(* IEC 61131-3 sources: Antarbhukti-LLM/DatasetCreation/SeedSTs/batch2_filtered_NETWORK (part 2) *)

(* ---- HTTP_GET.ST ---- *)
(*@PROPERTIES_EX@
TYPE: POU
LOCALE: 0
IEC_LANGUAGE: ST
PLC_TYPE: independent
PROC_TYPE: independent
GROUP: NETWORK
*)
(*@KEY@:DESCRIPTION*)

version 1.3	12. apr. 2011
programmer 	ks
tested by	ks

HTTP_GET führt eine HTTP Abfrage einer Web-Seite bei einem WEB_Server durch, und stellt die Daten ausbereitet zu verfügung
(*@KEY@:END_DESCRIPTION*)
FUNCTION_BLOCK HTTP_GET

(*Group:Default*)

VAR_IN_OUT
	URL_DATA :	oscat_url;
	IP_C :	oscat_IP_C;(*IP_Control Verwaltungsstruktur*)
	S_BUF :	oscat_NETWORK_BUFFER;
	R_BUF :	oscat_NETWORK_BUFFER;
END_VAR

VAR_INPUT
	IP4 :	DWORD;
	GET :	BOOL;
	MODE :	BYTE := BYTE#2;
	UNLOCK_BUF :	BOOL;
END_VAR

VAR_OUTPUT
	HTTP_STATUS :	STRING;
	HEADER_START :	UINT;(*HTTP Header (Message Header)*)
	HEADER_STOP :	UINT;(*HTTP Header (Message Header)*)
	BODY_START :	UINT;(*Message Body*)
	BODY_STOP :	UINT;(*Message Body*)
	DONE :	BOOL;
	ERROR :	DWORD;
END_VAR

VAR
	READ_HTTP :	READ_HTTP;
	BUFFER_SEARCH :	BUFFER_SEARCH_NW;
	_STRING_TO_BUFFER :	_STRING_TO_BUFFER_NW;
	IP_FIFO :	IP_FIFO;
	IS_NUM :	IS_NUM;
	ip_state :	BYTE;
	ip_id :	BYTE;
	get_last :	BOOL;
	ip4_stored :	DWORD;
	state :	INT;
	i :	INT;
	http_1_1_host :	BOOL;
	total_size :	INT;
	text :	oscat_STRING250;
	delimiter2b :	oscat_STRING2;
	delimiter4b :	oscat_STRING4;
	del_end :	oscat_STRING4;
	del_pos :	INT;
	idx :	INT;
	rcv_timeout :	BOOL;
	con_rdce :	BOOL;
END_VAR

(*Group:debug*)

VAR
	(*<LOG_MSG :	LOG_MSG;>*)
END_VAR

VAR_EXTERNAL
	(*<LOG_CL :	us_LOG_CONTROL;>*)(*Debug-Datenstruktur*)
END_VAR

VAR
	(*<_debug_enable :	BOOL := TRUE;>*)
END_VAR

(*@KEY@: WORKSHEET
NAME: HTTP_GET
IEC_LANGUAGE: ST
*)

CASE state OF
00:	IF GET AND NOT get_last THEN (* auf positive Flanke SET warten *)
		state        := 10;
		ip4_stored   := IP4; (* aktuelle IP4 speichern *)
		DONE         := FALSE;
		total_size   := 0;
		HEADER_START := UINT#0;
		HEADER_STOP  := UINT#0;
		BODY_START   := UINT#0;
		BODY_STOP    := UINT#0;
		HTTP_STATUS  := '';
    	ERROR        := DWORD#0;
    	ip_state     := BYTE#1; (* Anmelden *)

    	(* workaround für pcworx -> kein $0D$0A als Stringkonstante möglich *)
    	delimiter2b := CONCAT(BYTE_TO_STRING(BYTE#16#0D,'%c'),BYTE_TO_STRING(BYTE#16#0A,'%c'));
    	delimiter4b := CONCAT(delimiter2b,delimiter2b);
        (*####################  DEBUG-MESSAGE  ###################################*)
        (*IF _debug_enable THEN
            LOG_CL.NEW_MSG := 'HTTP: S00 START /IP_ID ~4';
            LOG_CL.PRINTF[4]  := BYTE_TO_STRING(IP_ID,'%u');
            LOG_MSG();
        END_IF;*)
        (*########################################################################*)
  	END_IF;

10:	IF ip_state = BYTE#3 THEN (* Bei IP_Control anmelden und auf freigabe warten *)
		idx := 0;
		text := CONCAT('GET ',URL_DATA.PATH);
		_STRING_TO_BUFFER(STR:=text,POS:=idx,PT:=S_BUF.BUFFER,SIZE:=UINT#4096); (* GET path in buffer kopieren *)
		S_BUF.BUFFER:=_STRING_TO_BUFFER.pt;
		idx := idx + LEN(text);

		IF LEN(URL_DATA.QUERY) > 0 THEN
			S_BUF.BUFFER[idx] := BYTE#63; (* ASCII '?' *)
			idx := idx + 1;
			_STRING_TO_BUFFER(STR:=URL_DATA.QUERY,POS:=idx,PT:=S_BUF.BUFFER,SIZE:=UINT#4096); (* QUERY in buffer kopieren *)
			S_BUF.BUFFER:=_STRING_TO_BUFFER.pt;
			idx := idx + LEN(URL_DATA.QUERY);
		END_IF;

		IF MODE >= BYTE#2 THEN (* gewünschte HTTP Version uebergeben *)
			text := ' HTTP/1.1';
		ELSE
			text := ' HTTP/1.0';
		END_IF;
		text := CONCAT(text,delimiter2b);
		_STRING_TO_BUFFER(STR:=text,POS:=idx,PT:=S_BUF.BUFFER,SIZE:=UINT#4096); (* HTTP Version in buffer kopieren *)
		S_BUF.BUFFER:=_STRING_TO_BUFFER.pt;
		idx := idx + LEN(text);

		IF MODE = BYTE#1 THEN (* HTTP/1.0 mit persistenter Verbindung gewünscht *)
			text := CONCAT('Connection: Keep-Alive',delimiter2b); (* workaround für pcworx -> kein $0D$0A als Stringkonstante möglich *)
		ELSIF MODE = BYTE#3 THEN (* HTTP/1.1 ohne persistenter Verbindung gewünscht *)
			text := CONCAT('Connection: Close',delimiter2b); (* workaround für pcworx -> kein $0D$0A als Stringkonstante möglich *)
		ELSE
			text := '';
		END_IF;
		text := CONCAT(text,URL_DATA.HEADER);
		_STRING_TO_BUFFER(STR:=text,POS:=idx,PT:=S_BUF.BUFFER,SIZE:=UINT#4096); (* HTTP Version in buffer kopieren *)
		S_BUF.BUFFER:=_STRING_TO_BUFFER.pt;
		idx := idx + LEN(text);

		text := CONCAT('Host: ',URL_DATA.DOMAIN);
		text := CONCAT(text,delimiter4b); (* workaround für pcworx -> kein $0D$0A als Stringkonstante möglich *)
		_STRING_TO_BUFFER(STR:=text,POS:=idx,PT:=S_BUF.BUFFER,SIZE:=UINT#4096); (* HTTP Host in buffer kopieren *)
		S_BUF.BUFFER:=_STRING_TO_BUFFER.pt;
		idx := idx + LEN(text);

		(* IP Datenverkehr einrichten *)
		IF URL_DATA.PORT = WORD#0 THEN
			IP_C.C_PORT    := WORD#80;        (* Standard-Portnummer verwenden               *)
		ELSE
			IP_C.C_PORT    := URL_DATA.PORT;  (* Portnummer aus URL verwenden                *)
		END_IF;

		IP_C.C_IP       := ip4_stored;       (* IP eintragen                                  *)
		IP_C.C_MODE     := BYTE#0;           (* Mode: TCP+AKTIV+PORT+IP                       *)
		IP_C.C_ENABLE   := TRUE;             (* Verbindungsaufbau freigeben                   *)
		IP_C.TIME_RESET := TRUE;             (* Zeitueberwachung rücksetzen                   *)
		IP_C.R_OBSERVE  := TRUE;             (* Datenempfang ueberwachen                      *)
		S_BUF.SIZE      := INT_TO_UINT(idx); (* Sendelänge eintragen                          *)
		R_BUF.SIZE      := UINT#0;           (* Empfangslänge rücksetzen                      *)

		state := 30;
        (*####################  DEBUG-MESSAGE  ###################################*)
        (*IF _debug_enable THEN
            LOG_CL.NEW_MSG := 'HTTP: S20 SEND /IP_ID ~4';
            LOG_CL.PRINTF[4]  := BYTE_TO_STRING(IP_ID,'%u');
            LOG_MSG();
        END_IF;*)
        (*########################################################################*)

	END_IF;

30:	rcv_timeout := (IP_C.ERROR AND DWORD#16#0000_FF00) = DWORD#16#0000_FF00;
	con_rdce := (IP_C.ERROR AND DWORD#16#FD00_0000) = DWORD#16#FD00_0000;

	IF S_BUF.SIZE = UINT#0 THEN
		IF total_size = 0 THEN
			IF R_BUF.SIZE > UINT#15 THEN;  (* länge der empfangenen Daten prüfen *)

				(* HTTP HEADER Ende suchen -> durch $0D$A$0D$A erkennbar bei DEC RT-11,CP/M,MS-DOS,Windows *)
				del_end := delimiter4b;

				BUFFER_SEARCH(size:=R_BUF.SIZE,str:=del_end,pos:=0,ign:=FALSE,pt:=R_BUF.BUFFER);
				R_BUF.BUFFER:=BUFFER_SEARCH.pt;
				del_pos := BUFFER_SEARCH.BUFFER_SEARCH;

				(* kein Ende gefunden ? -> andere Ende-Codierung suchen *)
				IF del_pos = 0 THEN
          			(* workaround für pcworx -> kein $0A$0A als Stringkonstante möglich *)
          			del_end := CONCAT(BYTE_TO_STRING(BYTE#16#0A,'%c'),BYTE_TO_STRING(BYTE#16#0A,'%c'));

          			(* HTTP HEADER Ende suchen -> durch $A$A erkennbar bei Multics, Unix-Derivate,Mac OS X *)
          			BUFFER_SEARCH(size:=R_BUF.SIZE,str:=del_end,pos:=0,ign:=FALSE,pt:=R_BUF.BUFFER);
          			R_BUF.BUFFER:=BUFFER_SEARCH.pt;
		  			del_pos := BUFFER_SEARCH.BUFFER_SEARCH;
        		END_IF;

				IF del_pos > 0 THEN
					HEADER_START := UINT#0;
					HEADER_STOP  := INT_TO_UINT(del_pos + LEN(del_end) - 1);
					TOTAL_SIZE   := -1; (* HTTP Header empfangen aber noch keine gesamtlänge bekannt *)
				END_IF;

                (*####################  DEBUG-MESSAGE  ###################################*)
                (*IF _debug_enable THEN
                    LOG_CL.NEW_MSG := 'HTTP: S20 HEADER_START ~1 / HEADER_STOP ~2/IP_ID ~4';
                    LOG_CL.PRINTF[4]  := BYTE_TO_STRING(IP_ID,'%u');
                    LOG_CL.PRINTF[1]  := UINT_TO_STRING(HEADER_START,'%u');
                    LOG_CL.PRINTF[2]  := UINT_TO_STRING(HEADER_STOP,'%u');
                    LOG_MSG();
                END_IF;*)
                (*########################################################################*)

				(* HTTP Statuscode auswerten: (kann 1.0 oder 1.1 sein *)
				READ_HTTP(size:=HEADER_STOP,pos:=0,SRC:='',pt:=R_BUF.BUFFER);
				R_BUF.BUFFER:=READ_HTTP.pt;

				i := LEN(READ_HTTP.READ_HTTP);
				IF i > 7 THEN
					(* HTTP Version von HOST auswerten 1.0 oder 1.1 *)
					text:=MID(READ_HTTP.READ_HTTP,1,3);
					http_1_1_host := EQ_STRING(text,'1');

					(* Code und Meldung isolieren *)
					HTTP_STATUS := RIGHT(READ_HTTP.READ_HTTP,i - 4);
				END_IF;

				(* positive HTTP Anfrage ? *)
				IF FIND(HTTP_STATUS,'200') > 0 THEN

					(* 'Content-Length: Wert einlesen auswerten *)
					READ_HTTP(size:=HEADER_STOP,pos:=0,SRC:='CONTENT-LENGTH',pt:=R_BUF.BUFFER);
					R_BUF.BUFFER:=READ_HTTP.pt;
					text:=READ_HTTP.READ_HTTP;

					IF LEN(text) > 0 AND LEN(text) <= 80 THEN
						IS_NUM(str:=text);
						IF IS_NUM.IS_NUM THEN
							(* erwartete gesamtmenge an Bytes berechnen *)
							total_size := STRING_TO_INT(text)+ UINT_TO_INT(HEADER_STOP) + 1;
                            (*####################  DEBUG-MESSAGE  ###################################*)
                            (*IF _debug_enable THEN
                                LOG_CL.NEW_MSG := 'HTTP: S20 HEADER ~1, BODY ~2 TOTAL ~3 /IP_ID ~4';
                                LOG_CL.PRINTF[4]  := BYTE_TO_STRING(IP_ID,'%u');
                                LOG_CL.PRINTF[1]  := UINT_TO_STRING(HEADER_STOP,'%u');
                                LOG_CL.PRINTF[2]  := INT_TO_STRING(TOTAL_SIZE-UINT_TO_INT(HEADER_STOP),'%d');
                                LOG_CL.PRINTF[3]  := INT_TO_STRING(TOTAL_SIZE,'%d');
                                LOG_MSG();
                            END_IF;*)
                            (*########################################################################*)
						END_IF;
					END_IF;
				ELSE
					ERROR := DWORD#16#000000FC; (* Fehler durch HTTP-Statuscodes *)
				END_IF;
			END_IF;
			(* 1. bei bekannter Content-Length wird nach erhalt der erwartenen Daten die verbindung beendet *)
			(* 2. bei persistenter Verbindung muss bei unbekannter Datenmenge auf Receive-Timeout gewartet werden *)
			(* 3. wenn nach datenempfang die verbindung vom host unterbrochen wird *)
		ELSIF (R_BUF.SIZE >= INT_TO_UINT(total_size)) OR
			(R_BUF.SIZE > UINT#0 AND total_size < 0 AND ((rcv_timeout OR con_rdce) OR (IP_C.C_STATE = BYTE#1))) THEN

			IF R_BUF.SIZE - UINT#1 > HEADER_STOP THEN (* BODY Daten vorhanden *)
				BODY_START := HEADER_STOP + UINT#1;
				BODY_STOP  := R_BUF.SIZE - UINT#1;
                (*####################  DEBUG-MESSAGE  ###################################*)
                (*IF _debug_enable THEN
                    LOG_CL.NEW_MSG := 'HTTP: S20 BODY ~1, START ~2 END ~3 /IP_ID ~4';
                    LOG_CL.PRINTF[4]  := BYTE_TO_STRING(IP_ID,'%u');
                    LOG_CL.PRINTF[1]  := UINT_TO_STRING(HEADER_STOP,'%u');
                    LOG_CL.PRINTF[2]  := UINT_TO_STRING(BODY_START,'%u');
                    LOG_CL.PRINTF[3]  := UINT_TO_STRING(BODY_STOP,'%u');
                    LOG_MSG();
                END_IF;*)
                (*########################################################################*)

			END_IF;

			DONE := TRUE;
			IP_C.C_ENABLE := FALSE; (* Verbindung abbauen  *)
			state := 40;
            (*####################  DEBUG-MESSAGE  ###################################*)
            (*IF _debug_enable THEN
                LOG_CL.NEW_MSG := 'HTTP: S30 OK /IP_ID ~4';
                LOG_CL.PRINTF[4]  := BYTE_TO_STRING(IP_ID,'%u');
                LOG_MSG();
            END_IF;*)
            (*########################################################################*)
		END_IF;
	END_IF;

	IF IP_C.ERROR <> DWORD#0 THEN
		(* bei unbekannter Content-size ist nicht bekannt ob bzw wieviele Telegramme noch folgen werden *)
		(* darum wird nach receive-timeout oder Remote disconnect error der fehler wieder ausgefiltert (logischer fehler) *)
		IF rcv_timeout AND DONE THEN
			IP_C.ERROR := IP_C.ERROR AND DWORD#16#FFFF_00FF; (* Fehler wieder rücksetzen *)
		ELSIF con_rdce AND DONE THEN
			IP_C.ERROR := IP_C.ERROR AND DWORD#16#00FF_FFFF; (* Fehler wieder rücksetzen *)
		ELSE
			ERROR := IP_C.ERROR;
		END_IF;
	END_IF;

	IF ERROR > DWORD#0 THEN
		IP_C.C_ENABLE := FALSE; (* Verbindungsaufbau sperren           *)
		state := 40;
        (*####################  DEBUG-MESSAGE  ###################################*)
        (*IF _debug_enable THEN
            LOG_CL.NEW_MSG := 'HTTP: S30 ERROR ~1 /IP_ID ~4';
            LOG_CL.PRINTF[1]  := DWORD_TO_STRING(ERROR,'%08X');
            LOG_CL.PRINTF[4]  := BYTE_TO_STRING(IP_ID,'%u');
            LOG_MSG();
        END_IF;*)
        (*########################################################################*)
	END_IF;

40:	IF (UNLOCK_BUF OR NOT DONE) THEN (* Warten auf Release und Verbindung beendet -> IP_ID vom Stack nehmen *)
		IP_STATE := BYTE#4; (* Abmelden *)
		DONE := FALSE;
		state := 0;
	END_IF;
END_CASE;

GET_LAST := GET; (* letzten Status sichern zur Flankenerkennung *)

(* IP_FIFO *)
IP_FIFO(FIFO:=IP_C.FIFO,STATE:=ip_state,ID:=ip_id);
IP_C.FIFO:=IP_FIFO.FIFO;
ip_state:=IP_FIFO.STATE;
ip_id:=IP_FIFO.ID;

(* revision history
ks	18. oct. 2008	rev 1.0
	original version

ks	20. oct. 2009	rev 1.1
	Fehler bei body-suche bei $0a$0a korrigiert,Codeoptimierung,
	new VAR del_pos , del_end (Networkbuffer und Buffer-funktionen auf Basis 0)

ks	28. oct. 2009	rev 1.2
	über url.header können zusätzliche header-infos übergeben werden

ks	12. apr. 2011	rev 1.3
	verbesserte fehlererkennung und fehlerkorrektur bei buffer_to_string
*)

(*@KEY@: END_WORKSHEET *)
END_FUNCTION_BLOCK

(* ---- IP2GEO.ST ---- *)
(*@PROPERTIES_EX@
TYPE: POU
LOCALE: 0
IEC_LANGUAGE: ST
PLC_TYPE: independent
PROC_TYPE: independent
GROUP: NETWORK
*)
(*@KEY@:DESCRIPTION*)

version 	1.1	07.oct. 2010
programmer 	ks
tested by	ks

IP2GEO ermittelt die aktuelle WAN-IP und die dazugehörigen geographischen Infos

zusatzinfos: http://www.worldtimezone.com/time/wtzresult.php?CiID=10182&forma=

example:

http://ipinfodb.com/ip_query.php?timezone=true&IP=

<?xml version="1.0" encoding="UTF-8" ?>
- <Response>
  <Ip>85.127.218.109</Ip>
  <Status>OK</Status>
  <CountryCode>AT</CountryCode>
  <CountryName>Austria</CountryName>
  <RegionCode>09</RegionCode>
  <RegionName>Wien</RegionName>
  <City>Vienna</City>
  <ZipPostalCode />
  <Latitude>48.2</Latitude>
  <Longitude>16.3667</Longitude>
  <TimezoneName>Europe/Vienna</TimezoneName>
  <Gmtoffset>7200</Gmtoffset>
  <Isdst>1</Isdst>
  </Response>

(*@KEY@:END_DESCRIPTION*)
FUNCTION_BLOCK IP2GEO

(*Group:in_out*)

VAR_IN_OUT
	IP_C :	oscat_IP_C;(*IP_Control Verwaltungsstruktur*)
	S_BUF :	oscat_NETWORK_BUFFER;
	R_BUF :	oscat_NETWORK_BUFFER;
	GEO :	oscat_IP2GEO_DATA;
END_VAR

VAR_INPUT
	IP :	DWORD;
	ACTIVATE :	BOOL;
END_VAR

VAR_OUTPUT
	BUSY :	BOOL;
	DONE :	BOOL;
	ERROR_C :	DWORD;
	ERROR_T :	BYTE;
END_VAR

(*Group:var*)

VAR
	CTRL :	oscat_XML_CONTROL;
	XML_READER :	XML_READER;
	URL_DATA :	oscat_url;
	DNS_CLIENT :	DNS_CLIENT;
	STRING_TO_URL :	STRING_TO_URL;
	HTTP_GET :	HTTP_GET;
	FLOAT_TO_REAL :	FLOAT_TO_REAL;
	last_state :	BOOL;
	value_int :	INT;
	value_real :	REAL;
	v_real :	REAL;
	state :	INT;
	IP4_TO_STRING :	IP4_TO_STRING;
	IP4_DECODE :	IP4_DECODE;
	CHK_REAL :	CHK_REAL;
END_VAR

(*@KEY@: WORKSHEET
NAME: IP2GEO
IEC_LANGUAGE: ST
*)

CASE state OF

00:
  IF ACTIVATE AND NOT last_state THEN
    state := 20;
	DONE := FALSE;
	BUSY := TRUE;
	ERROR_C := DWORD#0;
	ERROR_T := BYTE#0;
  END_IF;

20: (* URL for DNS UND HTTP-GET *)
  (* Example: http://ipinfodb.com/ip_query.php?timezone=true&IP=10.10.10.10 *)
  STRING_TO_URL.STR:='http://ipinfodb.com/ip_query.php?timezone=true&IP=';
  STRING_TO_URL.DEFAULT_PROTOCOL:='';
  STRING_TO_URL.DEFAULT_PATH:='';
  STRING_TO_URL();
  URL_DATA:=STRING_TO_URL.STRING_TO_URL;

  IF IP > DWORD#0 THEN
    IP4_TO_STRING(IP4:=IP);
    URL_DATA.QUERY := CONCAT(URL_DATA.QUERY,IP4_TO_STRING.IP4_TO_STRING);
  END_IF;

  state := 40;

40:
  IF DNS_CLIENT.DONE THEN
    state := 60;
  ELSIF (DNS_CLIENT.ERROR > DWORD#00) THEN
    (* Fehlerbehandlung *)
    ERROR_C := DNS_CLIENT.ERROR;
	ERROR_T := BYTE#01;
    state   := 100;
  END_IF;

60:
  IF HTTP_GET.DONE THEN
    state := 80;
    CTRL.START_POS := HTTP_GET.BODY_START;
    CTRL.STOP_POS  := HTTP_GET.BODY_STOP;
    CTRL.COMMAND   := WORD#2#10000000_00011000; (* ONLY TEXT AND ATTRIBUTE *)
	CTRL.WATCHDOG  := T#1ms;

  ELSIF (HTTP_GET.ERROR > DWORD#00) THEN
    (* Fehlerbehandlung *)
    ERROR_C := HTTP_GET.ERROR;
	  ERROR_T := BYTE#02;
    state   := 100;
  END_IF;

80:
  (* XML Daten seriell lesen *)
  XML_READER.CTRL := CTRL;
  XML_READER.BUF  := R_BUF.BUFFER;
  XML_READER();
  CTRL         := XML_READER.CTRL;
  R_BUF.BUFFER := XML_READER.BUF;

  IF CTRL.TYP < 98 THEN (* nur auswerten wenn kein Watchdog durchlauf *)
		(* automatische konvertierung in real und int ausführen *)
		value_int := 0;
		value_real := 0.0;
		IF LEN(CTRL.VALUE) <= 20 THEN
      		FLOAT_TO_REAL(FLT:=CTRL.VALUE);
			v_real :=FLOAT_TO_REAL.FLOAT_TO_REAL;
			CHK_REAL(X:= v_real); (* !!! prüft auf gültigen REAL Wert, ansonsten stürzt Twincat ab !!!!  *)
			IF CHK_REAL.CHK_REAL = BYTE#0 THEN
				value_real := v_real;
				value_int := REAL_TO_INT(value_real);
			END_IF;
		END_IF;

    CASE UINT_TO_INT(CTRL.COUNT) OF

      07: IP4_DECODE(STR:=CTRL.VALUE);
          GEO.IP4 := IP4_DECODE.IP4_DECODE; (* IP-Adresse *)
	  10: GEO.STATE := EQ_STRING('OK',CTRL.VALUE); (* STATUS *)
	  13: GEO.COUNTRY_CODE := CTRL.VALUE; (* Country-Code *)
	  16: GEO.COUNTRY_NAME := CTRL.VALUE; (* Country-Name *)
	  19: GEO.REGION_CODE := CTRL.VALUE; (* Region-Code *)
	  22: GEO.REGION_NAME := CTRL.VALUE; (* Region-Name *)
	  25: GEO.CITY := CTRL.VALUE; (* City *)
	  31: GEO.GEO_LATITUDE := value_real; (* Latitude *)
	  34: GEO.GEO_LONGITUDE := value_real; (* Longitude *)
	  37: GEO.TIME_ZONE_NAME := CTRL.VALUE; (* TimeZone Name *)
	  40: GEO.GMT_OFFSET := value_int; (* GMT OFFSET in Minuten *)
	  43: GEO.IS_DST := value_int > 0; (* Sommerzeit aktiv *)
    END_CASE;

  ELSIF CTRL.TYP = 99 THEN (* EXIT - letztes Element gelesen *)
    DONE  := TRUE;
    state := 100;
  END_IF;

100:
  (* UNLOCK HTTP DATA *)
  IF (NOT HTTP_GET.DONE) THEN
    state := 0;
    BUSY  := FALSE;
    DONE := ERROR_T = BYTE#0;
  END_IF;

END_CASE;

(* ---------------- DNS --------------- *)
DNS_CLIENT.IP_C     := IP_C;
DNS_CLIENT.S_BUF    := S_BUF;
DNS_CLIENT.R_BUF    := R_BUF;
DNS_CLIENT.DOMAIN   := URL_DATA.DOMAIN;
DNS_CLIENT.IP4_DNS  := DWORD#00;
DNS_CLIENT.ACTIVATE := state=40; (* DNS Start *)
DNS_CLIENT();
IP_C  := DNS_CLIENT.IP_C;
S_BUF := DNS_CLIENT.S_BUF;
R_BUF := DNS_CLIENT.R_BUF;

(* nicht oder nicht direkt verwendete Parameter *)
(* DWORD :=DNS_CLIENT.IP4;
   BOOL  :=DNS_CLIENT.DONE;
   BYTE  :=DNS_CLIENT.ERROR; *)
(* -------------------------------------*)

(* ------------- HTTP_GET --------------- *)

HTTP_GET.IP_C        := IP_C;
HTTP_GET.S_BUF       := S_BUF;
HTTP_GET.R_BUF       := R_BUF;
HTTP_GET.IP4         := DNS_CLIENT.IP4;
HTTP_GET.GET         := state=60;
HTTP_GET.MODE        := BYTE#2; (* HTTP 1.1 mit persistenter Verbindung *)
HTTP_GET.UNLOCK_BUF  := state=100;
HTTP_GET.URL_DATA    := URL_DATA;
HTTP_GET();
IP_C     := HTTP_GET.IP_C;
S_BUF    := HTTP_GET.S_BUF;
R_BUF    := HTTP_GET.R_BUF;
URL_DATA := HTTP_GET.URL_DATA;

(* nicht oder nicht direkt verwendete Parameter *)
(*STRING := HTTP_GET.HTTP_STATUS;
  UINT :=HTTP_GET.HEADER_START;
  UINT :=HTTP_GET.HEADER_STOP;
  UINT :=HTTP_GET.BODY_START;
  UINT :=HTTP_GET.BODY_STOP;
  BOOL :=HTTP_GET.DONE;
  BYTE :=HTTP_GET.ERROR;
*)
(* -------------------------------------*)

last_state := ACTIVATE;

(* revision history
ks	14. aug. 2009	rev 1.0
	original version

ks	07. oct. 2010	rev 1.1
	new url , ip2geo fields , REAL_CHECK
*)

(*@KEY@: END_WORKSHEET *)
END_FUNCTION_BLOCK

(* ---- IP_CONTROL.ST ---- *)
(*@PROPERTIES_EX@
TYPE: POU
LOCALE: 0
IEC_LANGUAGE: ST
PLC_TYPE: independent
PROC_TYPE: independent
GROUP: HARDWARE
*)
(*@KEY@:DESCRIPTION*)

version 1.8		26. july. 2011
programmer 		ks
tested by		ks

IP_CONTROL ist ein Wrapper-Baustein um eine Hersteller neutrale Schnittstelle zum Ethernet zu schaffen

(*@KEY@:END_DESCRIPTION*)
FUNCTION_BLOCK IP_CONTROL

(*Group:debug*)

VAR
	(*<debug_index :	INT;>*)(*test debug*)
	(*<debug_ID :	INT;>*)(*test debug*)
	(*<debug_lasterror :	DWORD;>*)(*test debug*)
	(*<debug_last_id :	INT := 255;>*)(*test debug*)
	(*<_debug_enable :	BOOL := TRUE;>*)
END_VAR

VAR_EXTERNAL
	(*<LOG_CL :	us_LOG_CONTROL;>*)(*Debug-Datenstruktur*)
END_VAR

VAR
	(*<LOG_MSG :	LOG_MSG;>*)(*Debug-Bausteininstanz*)
END_VAR

(*Group:instance*)

VAR
	T_PLC_MS :	T_PLC_MS;(*Bausteininstanz T_PLC_MS*)
	IP4_TO_STRING :	IP4_TO_STRING;(*Bausteininstanz*)
	FB_IP_CONNECT :	IP_CONNECT;(*Bausteininstanz IP_CONNECT*)
	FB_IP_URCV :	IP_URCV;(*Bausteininstanz IP_RECEIVE*)
	FB_IP_USEND :	IP_USEND;(*Bausteininstanz IP_SEND*)
END_VAR

(*Group:IN_OUT*)

VAR_INPUT
	IP :	DWORD;(*IP Adresse*)
	PORT :	WORD;(*Port Nummer*)
	TIME_OUT :	TIME;(*Ueberwachungszeit Connect / Send / Receive*)
END_VAR

VAR_IN_OUT
	IP_C :	oscat_IP_C;(*IP_Control Verwaltungsstruktur*)
	S_BUF :	oscat_NETWORK_BUFFER;(*Externer Sendbuffer*)
	R_BUF :	oscat_NETWORK_BUFFER;(*Externer Receivebuffer*)
END_VAR

(*Group:lokal*)

VAR
	C_TIME :	UDINT;(*CONNECT-Time (Zeit bei nicht vorhandener Verbindung)*)
	S_TIME :	UDINT;(*SEND-Time    (Zeit seit letzten Datensenden)*)
	R_TIME :	UDINT;(*RECEIVE-Time (Zeit seit letztem Datenempfang)*)
	C_ENABLE :	BOOL;(*CONNECT freigabe*)
	C_IP :	DWORD;(*Connect: aktuelle IP-Adresse*)
	C_PORT :	WORD;(*Connect: aktuelle Port-Nummer*)
	C_MODE :	BYTE;(*Connect: aktueller Mode UDP/TCP......*)
	C_ERROR :	BOOL;(*Connect Error vorhanden*)
	C_STATUS :	INT;(*Connect Status (Errorcode)*)
	C_ID :	INT;(*Connect ID für Send und Receive Baustein*)
	C_RECONNECT :	BOOL;(*Reconnect durchführen*)
	C_RECONNECT_COUNT :	INT;(*Reconnect zähler*)
	S_BUF_I :	oscat_NETWORK_BUFFER_SHORT;(*interner Sendbuffer*)
	S_TOTAL :	INT;(*Gesamtanzahl Bytes zum senden*)
	S_CUR_POS :	INT;(*aktuelle Sendeposition*)
	S_CUR_SIZE :	INT;(*aktuelle Sendegroesse*)
	S_MAX_SIZE :	INT := 1408;(*maximale Telegrammlänge fuer Senden*)
	S_START :	BOOL;(*Mode für IP_SEND Aufruf*)
	S_REQ :	BOOL;(*pos. Flanke Start Daten senden*)
	S_DONE :	BOOL;(*Senden ohne Fehler beendet*)
	S_ERROR :	BOOL;(*Sende Error vorhanden*)
	S_STATUS :	INT;(*Sende Status (Errorcodes)*)
	R_NDR :	BOOL;(*pos. Flanke wenn neue Daten empfangen wurden*)
	R_ERROR :	BOOL;(*Receive Error vorhanden*)
	R_STATUS :	INT;(*Receive Status (Errorcodes)*)
	R_BUF_I :	oscat_NETWORK_BUFFER_SHORT;(*Interner Receivebuffer*)
	R_COUNT :	INT;(*Receive Anzahl empfangener Bytes*)
	R_OFFSET :	INT;(*aktuelle Position in externen Receivebuffer*)
	R_E_MAX_SIZE :	INT := 4096;(*groesse des externen Empfangbuffers*)
	NEW_CONNECTION :	BOOL;(*Neue Verbindungsparameter vorhanden*)
	C_ENABLE_OLD :	BOOL;(*letzter Zustand von C_ENABLE für Flankenauswertung*)
	C_READY :	BOOL;(*Verbindung aufgebaut*)
	C_READY_OLD :	BOOL;(*letzter Zustand von C_READY für Flankenauswertung*)
	DELAY_STOP :	UDINT;(*PCWORX Workaround*)
	DELAY :	UDINT;(*PCWORX Workaround*)
	DELAY_VALUE :	UDINT;(*PCWORX Workaround*)
	C :	INT;(*temp*)
	C2 :	INT;(*temp*)
	C3 :	INT;(*temp*)
	CS :	STRING;(*Connect PARTNER STRING*)
	TX :	UDINT;(*letzter zeitwert*)
	ERROR_TIME :	UDINT;(*aktueller Timeout-Wert*)
	S_ACTIVE :	BOOL;(*Daten senden ist aktiv*)
	ERROR_CON :	BYTE;(*Error Connect*)
	ERROR_SND :	BYTE;(*Error Send*)
	ERROR_RCV :	BYTE;(*Error Receive*)
END_VAR

(*@KEY@: WORKSHEET
NAME: CONNECT
IEC_LANGUAGE: ST
*)
(* read system time *)
T_PLC_MS();
TX := T_PLC_MS.T_PLC_MS;

(*++++++ PCWORX spez. Sonderbehandlung bei Connect on/off ++++++++++++++++++*)

(* bei Connect on/off aktivitäten muss die abarbeitung zeitverzögert werden *)
IF (TX - DELAY < DELAY_VALUE) THEN
  IF IP_C.C_STATE <> BYTE#1 AND IP_C.C_STATE <> BYTE#254 THEN (* Bei vorhandenen Connect OFF/ON Flankenmeldungen die abarbeitet nicht unterbrechen *)
	RETURN;
  END_IF;
END_IF;
DELAY := TX;

(*####################  DEBUG-MESSAGE  ###################################*)
(*IF _debug_enable THEN
	IF IP_C.FIFO.ID > BYTE#0 THEN
		debug_index := IP_C.FIFO.NR;
    	debug_ID := BYTE_TO_INT(IP_C.FIFO.X[debug_index]);
	END_IF;
END_IF;*)
(*########################################################################*)

(* Connect on/off verzoegerung nach 1000ms wieder zurücknehmen *)
IF C_ENABLE AND DELAY_VALUE > UDINT#00 THEN
  IF (TX - DELAY_STOP > UDINT#1000) THEN
    DELAY_VALUE := UDINT#00;
    (*####################  DEBUG-MESSAGE  ###################################*)
    (*IF _debug_enable THEN
      LOG_CL.NEW_MSG := 'IP_CON: STOP CYCLE_DELAY -IP_ID ~6';
      LOG_CL.PRINTF[1] := CS;
      LOG_CL.PRINTF[6] := INT_TO_STRING(debug_ID,'%d');
      LOG_MSG();
    END_IF;*)
    (*########################################################################*)
  END_IF;
ELSE
  DELAY_STOP := TX;  (* timer starten              *)
END_IF;
(*++++++++++++++++++++++++++++++++++++++++++++++++++++++++++++++++++++++++++*)

(* -----------------------------------------------------------------*)
(* wenn ein satelliten-baustein die portnummer 0 oder IP-Adresse    *)
(* 0.0.0.0 verwendet, sollen die am ip_control angegebene daten     *)
(* verwendet werden.           										*)
(* -----------------------------------------------------------------*)
IF IP_C.C_PORT = WORD#00 THEN
	IP_C.C_PORT := PORT; (* uebergebenen PORT durch paramtrierte PORT ersetzen *)
END_IF;
IF IP_C.C_IP=DWORD#00 AND IP_C.C_MODE<BYTE#4 THEN
	IP_C.C_IP := IP; (* uebergebene IP durch paramtrierte IP ersetzen *)
END_IF;

(* neue Verbindungs erwünscht ? *)
NEW_CONNECTION := C_IP <> IP_C.C_IP OR C_MODE <> IP_C.C_MODE OR C_PORT <> IP_C.C_PORT;

(* -----------------------------------------------------------------*)
(* Verbindungsparameter ausbereiten                                 *)
(* -----------------------------------------------------------------*)
IF IP_C.C_ENABLE AND NOT C_READY AND NEW_CONNECTION THEN

  (* neue Verbindungsparameter übernehmen *)
  C_IP   := IP_C.C_IP;
  C_MODE := IP_C.C_MODE;
  C_PORT := IP_C.C_PORT;

  (* -----------------------------------------------------------------*)
  (* CONNECTION_STRING erzeugen                                       *)
  (* Beispiel: '/UDP /ACTIVE /PORT=1000 /IP=192.168.178.1'            *)
  (*                                                                  *)
  (* Mode:                                                            *)
  (*  0: TCP + ACTIVE  + PORT + IP                                    *)
  (*  1: UDP + ACTIVE  + PORT + IP                                    *)
  (*  2: TCP + PASSIVE + PORT + IP                                    *)
  (*  3: UDP + PASSIVE + PORT + IP                                    *)
  (*  4: TCP + PASSIVE + PORT                                         *)
  (*  5: UDP + PASSIVE + PORT                                         *)
  (* -----------------------------------------------------------------*)

  (* bei allen ungeraden MODE Nummern UDP-String vorgeben *)
  CS := SEL_STRING((C_MODE AND BYTE#1) = BYTE#1,'','/UDP');
  (* ACTIVE oder PASSIVE String anhängen *)
  CS := CONCAT(CS,SEL_STRING(C_MODE<BYTE#2,' /PASSIVE',' /ACTIVE'));
  (* Portnummer String anhängen *)
  CS := CONCAT(CS,' /PORT=');
  CS := CONCAT(CS,WORD_TO_STRING(C_PORT,'%u'));

  IF C_MODE<BYTE#4 THEN
    IP4_TO_STRING(IP4:=C_IP);  (* String mit IP erzeugen *)
    CS := CONCAT(CS,' /IP=');
    CS := CONCAT(CS,IP4_TO_STRING.IP4_TO_STRING);
  END_IF;

  (*-------------------------------------------------------------------*)

  (* uebergebenen Timeout-Wert auf min-wert begrenzen *)
  ERROR_TIME := MAX(UDINT#200,TIME_TO_UDINT(TIME_OUT));
  IP_C.TIME_RESET := TRUE;   (* Alle Timer ruecksetzen *)
  (*####################  DEBUG-MESSAGE  ###################################*)
  (*IF _debug_enable THEN
    LOG_CL.NEW_MSG := 'IP_CON: ~1 -IP_ID ~6';
    LOG_CL.PRINTF[1] := CS;
    LOG_CL.PRINTF[6] := INT_TO_STRING(debug_ID,'%d');
    LOG_MSG();
  END_IF;*)
  (*########################################################################*)

END_IF;

(*++++++++++++++++++++++++++++++++++++++++++++++++++++++++++++++++++++++++++*)

C_ENABLE := IP_C.C_ENABLE AND NOT C_RECONNECT AND NOT NEW_CONNECTION AND IP_C.ERROR = DWORD#0;

(* -----------------------------------------------------------------*)
(* Systembaustein IP_CONNECT                                        *)
(* -----------------------------------------------------------------*)
FB_IP_CONNECT.EN_C    := C_ENABLE;
FB_IP_CONNECT.PARTNER := CS;
FB_IP_CONNECT();
C_READY  := FB_IP_CONNECT.VALID;
C_ERROR  := FB_IP_CONNECT.ERROR;
C_STATUS := FB_IP_CONNECT.STATUS;
C_ID     := FB_IP_CONNECT.ID;

(*++++++++++++++++++++++++++++++++++++++++++++++++++++++++++++++++++++++++++*)

IF C_ENABLE THEN
  IF NOT C_ENABLE_OLD THEN
    DELAY_VALUE := UDINT#50;  (* verzoegerungzeit 50ms vorgeben               *)
    (*####################  DEBUG-MESSAGE  ###################################*)
    (*IF _debug_enable THEN
      LOG_CL.NEW_MSG := 'IP_CON: ENABLE + CYLCE-DELAY -IP_ID ~6';
      LOG_CL.PRINTF[6] := INT_TO_STRING(debug_ID,'%d');
      LOG_MSG();
    END_IF;*)
    (*########################################################################*)
  END_IF;
ELSE
  IF C_ENABLE_OLD THEN
    C_RECONNECT := FALSE;
    DELAY_VALUE := UDINT#50; (* verzoegerungzeit 50ms vorgeben                *)
    (*####################  DEBUG-MESSAGE  ###################################*)
    (*IF _debug_enable THEN
      LOG_CL.NEW_MSG := 'IP_CON: DISABLE + CYLCE-DELAY -IP_ID ~6';
      LOG_CL.PRINTF[6] := INT_TO_STRING(debug_ID,'%d');
      LOG_MSG();
    END_IF;*)
    (*########################################################################*)
  END_IF;
END_IF;

C_ENABLE_OLD := C_ENABLE;

(*++++++++++++++++++++++++++++++++++++++++++++++++++++++++++++++++++++++++++*)

IF C_READY THEN
  IF NOT C_READY_OLD THEN
    (* Verbindung aufgebaut - positive Flanke erkannt*)
    IP_C.C_STATE := BYTE#254;
    DELAY_VALUE := UDINT#50;  (* verzoegerungzeit 50ms vorgeben *)
    IP_C.TIME_RESET := TRUE;  (* Alle Timer ruecksetzen *)
    (*####################  DEBUG-MESSAGE  ###################################*)
    (*IF _debug_enable THEN
      LOG_CL.NEW_MSG := 'IP_CON: CONNECTED -IP_ID ~6';
      LOG_CL.PRINTF[6] := INT_TO_STRING(debug_ID,'%d');
      LOG_MSG();
    END_IF;*)
    (*########################################################################*)

  ELSE
    IP_C.C_STATE := BYTE#255;  (* Verbindung ist aufgebaut                      *)
  END_IF;
ELSE
  IF C_READY_OLD THEN
    (* Verbindung abgebaut - negative Flanke erkannt*)
    IP_C.C_STATE := BYTE#1;
	IP_C.MAILBOX[1] := BYTE#0; (* Receive Info rücksetzen *)
	IP_C.MAILBOX[2] := BYTE#0; (* Send-Pause rücksetzen *)
	IP_C.MAILBOX[3] := BYTE#0; (* Receive-Pause rücksetzen *)
    DELAY_VALUE := UDINT#50;  (* verzoegerungzeit 50ms vorgeben *)

    IF NOT NEW_CONNECTION THEN
      S_ACTIVE := FALSE;        (* Sendeaktivitäten stoppen *)
      S_REQ := FALSE;           (* Sendefreigabe rücksetzen *)
      S_BUF.SIZE := UINT#0;     (* Sendelänge löschen       *)
      (*IP_C.TIME_RESET := TRUE;*)  (* Alle Timer ruecksetzen   *)
    END_IF;
    (*####################  DEBUG-MESSAGE  ###################################*)
    (*IF _debug_enable THEN
      LOG_CL.NEW_MSG := 'IP_CON: DISCONNECTED';
      LOG_MSG();
    END_IF;*)
    (*########################################################################*)
  ELSE
    IP_C.C_STATE := BYTE#000; (* Verbindung ist abgebaut *)
  END_IF;
END_IF;

C_READY_OLD := C_READY;

(*++++++++++++++++++++++++++++++++++++++++++++++++++++++++++++++++++++++++++*)
(*@KEY@: END_WORKSHEET *)
(*@KEY@: WORKSHEET
NAME: SEND
IEC_LANGUAGE: ST
*)
C := 1; (* voreinstellung: USEND einmal durchlaufen *)
IF S_BUF.SIZE > UINT#0 THEN
  IF C_READY AND C_ENABLE THEN
    IF S_ACTIVE = FALSE AND IP_C.MAILBOX[2] = BYTE#0 THEN
	  (* Gesamtanzahl an Bytes limitieren und uebergeben *)
      S_TOTAL := LIMIT_INT(0,UINT_TO_INT(S_BUF.SIZE),R_E_MAX_SIZE);
      S_CUR_POS  := 0;
      S_CUR_SIZE := 0;
      S_START := TRUE;      (* Daten kopieren und senden anstossen *)
      S_ACTIVE := TRUE;     (* Sende-Betrieb aktivieren *)
      (*####################  DEBUG-MESSAGE  ###################################*)
      (*IF _debug_enable THEN
        LOG_CL.NEW_MSG := 'IP_SEN INIT: TOTAL: ~1 -IP_ID ~6';
        LOG_CL.PRINTF[1] := INT_TO_STRING(S_TOTAL,'%d');
        LOG_CL.PRINTF[6] := INT_TO_STRING(debug_ID,'%d');
        LOG_MSG();
      END_IF;*)
      (*########################################################################*)
    END_IF;

    (* Daten senden gewünscht *)
    IF S_DONE OR S_START THEN

      S_START := FALSE;
      S_CUR_POS := S_CUR_POS + S_CUR_SIZE;              (* neue Sende-Datenposition bestimmen *)
      IF S_TOTAL > S_CUR_POS THEN                      (* weitere Daten zum senden vorhanden ? *)
        S_CUR_SIZE := S_TOTAL - S_CUR_POS;
        S_CUR_SIZE:=LIMIT_INT(0,S_CUR_SIZE,S_MAX_SIZE); (* Telegrammlänge begrenzen *)

  	    C2 := S_CUR_POS;
		C3 := S_CUR_SIZE - 1;
		FOR C := 0 TO C3 DO (* Datacopy routine *)
          S_BUF_I.BUFFER[C] := S_BUF.BUFFER[C2];
		  C2 := C2 + 1;
        END_FOR;

        (*####################  DEBUG-MESSAGE  ###################################*)
        (*IF _debug_enable THEN
          LOG_CL.NEW_MSG := 'IP_SEN DATA: POS: ~1 : SIZE: ~2 TOTAL ~3 -IP_ID ~6';
          LOG_CL.PRINTF[1] := INT_TO_STRING(S_CUR_POS,'%d');
          LOG_CL.PRINTF[2] := INT_TO_STRING(S_CUR_SIZE,'%d');
          LOG_CL.PRINTF[3] := INT_TO_STRING(S_TOTAL,'%d');
          LOG_CL.PRINTF[6] := INT_TO_STRING(debug_ID,'%d');
          LOG_MSG();
        END_IF;*)
        (*########################################################################*)

        (* Sendelänge in Telegramm eintragen *)
        S_BUF_I.SIZE := INT_TO_UINT(S_CUR_SIZE);
	    S_TIME := tx; (* Send Timer ruecksetzen      *)
        R_TIME := tx; (* Receive Timer ruecksetzen *)
        S_REQ := TRUE;
        C := 0; (* USEND zweimal aufrufen zur erzeugung einer positiven Flanke *)

      ELSE
        (* keine weitere Sendedaten vorhanden -> Senden beenden *)
        S_REQ := FALSE;
        S_BUF.SIZE := UINT#0;
        S_ACTIVE := FALSE;
        (*####################  DEBUG-MESSAGE  ###################################*)
        (*IF _debug_enable THEN
          LOG_CL.NEW_MSG := 'IP_SEN FINISH -IP_ID ~6';
          LOG_CL.PRINTF[6] := INT_TO_STRING(debug_ID,'%d');
          LOG_MSG();
        END_IF;*)
        (*########################################################################*)
      END_IF;
    END_IF;
  END_IF;
END_IF;

(* -----------------------------------------------------------------*)
(* Systembaustein IP_USEND (Datensenden)                            *)
(* -----------------------------------------------------------------*)
FOR C2 := C TO 1 DO
  FB_IP_USEND.REQ    := S_REQ AND C2=1;
  FB_IP_USEND.ID     := C_ID;
  FB_IP_USEND.R_ID   := '';
  FB_IP_USEND.SD_1   := S_BUF_I;
  FB_IP_USEND();
  S_DONE   := FB_IP_USEND.DONE;
  S_ERROR  := FB_IP_USEND.ERROR;
  S_STATUS := FB_IP_USEND.STATUS;
  S_BUF_I  := FB_IP_USEND.SD_1;
END_FOR;
(*@KEY@: END_WORKSHEET *)
(*@KEY@: WORKSHEET
NAME: RECEIVE
IEC_LANGUAGE: ST
*)
(* -----------------------------------------------------------------*)
(* Systembaustein IP_URCV (Datenempfang)                            *)
(* -----------------------------------------------------------------*)
FB_IP_URCV.EN_R := C_READY AND NOT S_ACTIVE AND IP_C.MAILBOX[3] = BYTE#0;
FB_IP_URCV.ID   := C_ID;
FB_IP_URCV.R_ID := '';
FB_IP_URCV.RD_1 := R_BUF_I;
FB_IP_URCV();
R_NDR    := FB_IP_URCV.NDR;
R_ERROR  := FB_IP_URCV.ERROR;
R_STATUS := FB_IP_URCV.STATUS;
R_BUF_I  := FB_IP_URCV.RD_1;

(* -----------------------------------------------------------------*)
(* positive Flanke für Daten Empfangen abfragen                     *)
(* -----------------------------------------------------------------*)
IF R_NDR THEN
  IF R_BUF.SIZE >= INT_TO_UINT(R_E_MAX_SIZE) THEN
    R_BUF.SIZE := UINT#0;
    r_status := 254; (* Empfangsbuffer wegen Überlauf rückgesetzt *)
  END_IF;

  R_TIME := tx; (* Receive Timer ruecksetzen           *)
  R_COUNT := UINT_TO_INT(R_BUF_I.SIZE); (* Anzahl empfangener Bytes bestimmen *)
  R_OFFSET := UINT_TO_INT(R_BUF.SIZE); (* Start Offset Zielbuffer *)

  IF (C_MODE AND BYTE#2#0000_0001) = BYTE#1 THEN (* UDP MODE *)
    r_offset := 0; (* Daten immer ab position 0 ablegen -> kein Datastream *)
  ELSE
    R_OFFSET := UINT_TO_INT(R_BUF.SIZE); (* Start Offset Zielbuffer *)
  END_IF;

  (* Datenempfang auf buffergroesse beschränken *)
  IF R_OFFSET + R_COUNT > R_E_MAX_SIZE THEN
    R_COUNT := R_E_MAX_SIZE - R_OFFSET;
  END_IF;

  (* Datacopy routine *)
  C2 := R_OFFSET;
  C3 := R_COUNT - 1;
  FOR C := 0 TO C3 DO
    R_BUF.BUFFER[C2] := R_BUF_I.BUFFER[C];
    C2 := C2 + 1;
  END_FOR;

  R_BUF.SIZE := INT_TO_UINT(R_OFFSET + R_COUNT); (* aktuelle buffersize eintragen *)
  IP_C.MAILBOX[1] := USINT_TO_BYTE(BYTE_TO_USINT(IP_C.MAILBOX[1]) + USINT#1); (* Receive Info *)
  IF IP_C.MAILBOX[1] = BYTE#0 THEN IP_C.MAILBOX[1] := BYTE#1; END_IF;

  (*####################  DEBUG-MESSAGE  ###################################*)
  (*IF _debug_enable THEN
    LOG_CL.NEW_MSG := 'IP_REC DATA: POS: ~1 : SIZE: ~2 TOTAL ~3 -IP_ID ~6';
    LOG_CL.PRINTF[1] := INT_TO_STRING(R_OFFSET,'%d');
    LOG_CL.PRINTF[2] := INT_TO_STRING(R_COUNT,'%d');
    LOG_CL.PRINTF[3] := UINT_TO_STRING(R_BUF.SIZE,'%u');
    LOG_CL.PRINTF[6] := INT_TO_STRING(debug_ID,'%d');
    LOG_MSG();
  END_IF;*)
  (*########################################################################*)

END_IF;
(*@KEY@: END_WORKSHEET *)
(*@KEY@: WORKSHEET
NAME: ERROR
IEC_LANGUAGE: ST
*)
(* ----------------------------------------------------------------------------*)
(* Timer bearbeitung                                                           *)
(* ----------------------------------------------------------------------------*)
IF IP_C.TIME_RESET THEN     (* Alle Timer ruecksetzen      *)
  IP_C.TIME_RESET := FALSE; (* Reset rücksetzen            *)
  C_RECONNECT_COUNT := 0;   (* Reconnect zähler rücksetzen *)
  C_TIME := tx;             (* Connect   Timer ruecksetzen *)
  S_TIME := tx;             (* Send      Timer ruecksetzen *)
  R_TIME := tx;             (* Receive   Timer ruecksetzen *)

  ERROR_CON := BYTE#0;		(* Error Connect rücksetzen    *)
  ERROR_SND := BYTE#0;		(* Error Send rücksetzen       *)
  ERROR_RCV := BYTE#0;		(* Error Receive rücksetzen    *)
END_IF;

IF IP_C.R_OBSERVE = FALSE OR s_active THEN
    R_TIME := tx;
END_IF;

C_RECONNECT := FALSE;

(* ----------------------------------------------------------------------------*)
(* Error bearbeitung                                                           *)
(*                                                                             *)
(* bei pcworx ist nur wenn error = 1  der wert von status ein echter fehler    *)
(* status bekommt bei error "0" auch manchmal andere werte                     *)
(* ----------------------------------------------------------------------------*)

(* CONNECT Fehlercodes *)
IF ERROR_CON = BYTE#0 THEN
  IF C_ERROR THEN (* Die Verbindung wurde abgebrochen ignorieren *)
	IF C_STATUS = 16#31 THEN (* Die Verbindung wurde abgebrochen *)
		ERROR_CON := BYTE#253;
	ELSE
		ERROR_CON := INT_TO_BYTE(C_STATUS);
	END_IF;
  ELSIF TX - C_TIME > ERROR_TIME AND C_ENABLE AND NOT C_READY AND C_MODE < BYTE#2 THEN (* Connect Timeout *)
    IF C_RECONNECT_COUNT >= 3 THEN
      ERROR_CON := BYTE#255; (* Timeout-Fehler ausgeben *)
    ELSE
      C_TIME := TX; (* Connect   Timer ruecksetzen            *)
      C_RECONNECT_COUNT := C_RECONNECT_COUNT + 1;
      C_RECONNECT := TRUE;
      (*####################  DEBUG-MESSAGE  ###################################*)
      (*IF _debug_enable THEN
        LOG_CL.NEW_MSG := 'IP_CON: RECONNECT -IP_ID ~6';
        LOG_CL.PRINTF[6] := INT_TO_STRING(debug_ID,'%d');
        LOG_MSG();
      END_IF;*)
      (*########################################################################*)

    END_IF;
  END_IF;
END_IF;

(* SEND Fehlercodes *)
IF ERROR_SND = BYTE#0 THEN
  IF S_ERROR AND S_STATUS <> 16#65 THEN (* andere Bausteininstanz arbeitet mit dieser Verbindung *)
  	ERROR_SND := INT_TO_BYTE(S_STATUS);
  ELSIF TX - S_TIME > ERROR_TIME AND S_ACTIVE THEN (* Send Timeout *)
    ERROR_SND := BYTE#255; (* Timeout-Fehler ausgeben *)
  END_IF;
END_IF;

(* RECEIVE Fehlercodes *)
IF ERROR_RCV = BYTE#0 THEN
  IF R_ERROR AND (R_STATUS <> 16#33) AND (R_STATUS <> 16#31) AND (R_STATUS <> 16#65) THEN (* Receive Timeout,Verbindungsabbruch,andere Bausteininstanz arbeitet mit dieser Verbindung, ignorieren *)
  	ERROR_RCV := INT_TO_BYTE(R_STATUS);
  ELSIF TX - R_TIME > ERROR_TIME AND C_READY AND IP_C.R_OBSERVE THEN (* Receive Timeout *)
    ERROR_RCV := BYTE#255; (* Timeout-Fehler ausgeben *)
  END_IF;
END_IF;

IP_C.ERROR := DWORD_OF_BYTE(ERROR_CON,ERROR_SND,ERROR_RCV,BYTE#0);

(*####################  DEBUG-MESSAGE  ###################################*)
(*IF _debug_enable THEN
  IF (debug_last_id <> debug_ID) AND (IP_C.ERROR <> debug_lasterror) AND (IP_C.ERROR <> DWORD#00) THEN
    LOG_CL.NEW_MSG := 'IP_ERROR ~1 -IP_ID ~6';
    LOG_CL.PRINTF[1] := DWORD_TO_STRING(IP_C.ERROR,'%08X');
    LOG_CL.PRINTF[6] := INT_TO_STRING(debug_ID,'%d');
    LOG_MSG();
	debug_lasterror := IP_C.ERROR;
	debug_last_id   := debug_ID;
  END_IF;
END_IF;*)
(*########################################################################*)

(* revision history
ks	18. oct. 2008	rev 1.0
	original version
ks	05. jan. 2009	rev 1.1
	zusätzlichen Parameter "Port" hinzugefügt, und Code bei Verbindungsaufbau angepasst
ks	28. feb. 2009	rev 1.2
	connect code angepasst und verkürzung der zyklen bei Send
ks	20. oct. 2009	rev 1.3
	network_buffer basis 0
ks	06. dec. 2009	rev 1.4
	receive_count MAILBOX[1]
ks	10. nov. 2010	rev 1.5
	send_pause MAILBOX[2] and receive_pause MAILBOX[3]
ks	07. feb. 2011	rev 1.6
	Fehlercode 253 bei Remote-Verbindungsabbruch
ks	30. may. 2011	rev 1.7
	Fehler bei Empfangüberwachung
ks	26. jul. 2011	rev 1.8
	optimierung der Empfangsüberwachung
*)

(*@KEY@: END_WORKSHEET *)
END_FUNCTION_BLOCK

(* ---- IP_CONTROL2.ST ---- *)
(*@PROPERTIES_EX@
TYPE: POU
LOCALE: 0
IEC_LANGUAGE: ST
PLC_TYPE: independent
PROC_TYPE: independent
GROUP: HARDWARE
*)
(*@KEY@:DESCRIPTION*)

version 1.8		26. july. 2011
programmer 		ks
tested by		ks

IP_CONTROL ist ein Wrapper-Baustein um eine Hersteller neutrale Schnittstelle zum Ethernet zu schaffen

(*@KEY@:END_DESCRIPTION*)
FUNCTION_BLOCK IP_CONTROL2

(*Group:debug*)

VAR
	(*<debug_index :	INT;>*)(*test debug*)
	(*<debug_ID :	INT;>*)(*test debug*)
	(*<debug_lasterror :	DWORD;>*)(*test debug*)
	(*<debug_last_id :	INT := 255;>*)(*test debug*)
	(*<_debug_enable :	BOOL := TRUE;>*)
END_VAR

VAR_EXTERNAL
	(*<LOG_CL :	us_LOG_CONTROL;>*)(*Debug-Datenstruktur*)
END_VAR

VAR
	(*<LOG_MSG :	LOG_MSG;>*)(*Debug-Bausteininstanz*)
END_VAR

(*Group:instance*)

VAR
	T_PLC_MS :	T_PLC_MS;(*Bausteininstanz T_PLC_MS*)
	IP4_TO_STRING :	IP4_TO_STRING;(*Bausteininstanz*)
	FB_IP_CONNECT :	IP_CONNECT;(*Bausteininstanz IP_CONNECT*)
	FB_IP_URCV :	IP_URCV;(*Bausteininstanz IP_RECEIVE*)
	FB_IP_USEND :	IP_USEND;(*Bausteininstanz IP_SEND*)
END_VAR

(*Group:IN_OUT*)

VAR_INPUT
	IP :	DWORD;(*IP Adresse*)
	PORT :	WORD;(*Port Nummer*)
	TIME_OUT :	TIME;(*Ueberwachungszeit Connect / Send / Receive*)
END_VAR

VAR_IN_OUT
	IP_C :	oscat_IP_C;(*IP_Control Verwaltungsstruktur*)
	S_BUF :	oscat_NETWORK_BUFFER_SHORT;(*Externer Sendbuffer*)
	R_BUF :	oscat_NETWORK_BUFFER_SHORT;(*Externer Receivebuffer*)
END_VAR

(*Group:lokal*)

VAR
	C_TIME :	UDINT;(*CONNECT-Time (Zeit bei nicht vorhandener Verbindung)*)
	S_TIME :	UDINT;(*SEND-Time    (Zeit seit letzten Datensenden)*)
	R_TIME :	UDINT;(*RECEIVE-Time (Zeit seit letztem Datenempfang)*)
	C_ENABLE :	BOOL;(*CONNECT freigabe*)
	C_IP :	DWORD;(*Connect: aktuelle IP-Adresse*)
	C_PORT :	WORD;(*Connect: aktuelle Port-Nummer*)
	C_MODE :	BYTE;(*Connect: aktueller Mode UDP/TCP......*)
	C_ERROR :	BOOL;(*Connect Error vorhanden*)
	C_STATUS :	INT;(*Connect Status (Errorcode)*)
	C_ID :	INT;(*Connect ID für Send und Receive Baustein*)
	C_RECONNECT :	BOOL;(*Reconnect durchführen*)
	C_RECONNECT_COUNT :	INT;(*Reconnect zähler*)
	S_DONE :	BOOL;(*Senden ohne Fehler beendet*)
	S_ERROR :	BOOL;(*Sende Error vorhanden*)
	S_STATUS :	INT;(*Sende Status (Errorcodes)*)
	S_ACTIVE :	BOOL;(*Daten senden ist aktiv*)
	R_NDR :	BOOL;(*pos. Flanke wenn neue Daten empfangen wurden*)
	R_ERROR :	BOOL;(*Receive Error vorhanden*)
	R_STATUS :	INT;(*Receive Status (Errorcodes)*)
	NEW_CONNECTION :	BOOL;(*Neue Verbindungsparameter vorhanden*)
	C_ENABLE_OLD :	BOOL;(*letzter Zustand von C_ENABLE für Flankenauswertung*)
	C_READY :	BOOL;(*Verbindung aufgebaut*)
	C_READY_OLD :	BOOL;(*letzter Zustand von C_READY für Flankenauswertung*)
	DELAY_STOP :	UDINT;
	DELAY :	UDINT;
	DELAY_VALUE :	UDINT;
	C :	INT;(*temp*)
	C2 :	INT;(*temp*)
	CS :	oscat_STRING50;(*Connect PARTNER STRING*)
	TX :	UDINT;(*letzter zeitwert*)
	ERROR_TIME :	UDINT;(*aktueller Timeout-Wert*)
	ERROR_CON :	BYTE;(*Error Connect*)
	ERROR_SND :	BYTE;(*Error Send*)
	ERROR_RCV :	BYTE;(*Error Receive*)
END_VAR

(*@KEY@: WORKSHEET
NAME: CONNECT
IEC_LANGUAGE: ST
*)
(* read system time *)
T_PLC_MS();
TX := T_PLC_MS.T_PLC_MS;

(*++++++ PCWORX spez. Sonderbehandlung bei Connect on/off ++++++++++++++++++*)

(* bei Connect on/off aktivitäten muss die abarbeitung zeitverzögert werden *)
IF (TX - DELAY < DELAY_VALUE) THEN
  IF IP_C.C_STATE <> BYTE#1 AND IP_C.C_STATE <> BYTE#254 THEN (* Bei vorhandenen Connect OFF/ON Flankenmeldungen die abarbeitet nicht unterbrechen *)
	RETURN;
  END_IF;
END_IF;
DELAY := TX;

(*####################  DEBUG-MESSAGE  ###################################*)
(*IF _debug_enable THEN
	IF IP_C.FIFO.ID > BYTE#0 THEN
		debug_index := IP_C.FIFO.NR;
    	debug_ID := BYTE_TO_INT(IP_C.FIFO.X[debug_index]);
	END_IF;
END_IF;*)
(*########################################################################*)

(* Connect on/off verzoegerung nach 1000ms wieder zurücknehmen *)
IF C_ENABLE AND DELAY_VALUE > UDINT#00 THEN
  IF (TX - DELAY_STOP > UDINT#1000) THEN
    DELAY_VALUE := UDINT#00;
    (*####################  DEBUG-MESSAGE  ###################################*)
    (*IF _debug_enable THEN
      LOG_CL.NEW_MSG := 'IP_CON: STOP CYCLE_DELAY -IP_ID ~6';
      LOG_CL.PRINTF[1]  := CS;
      LOG_CL.PRINTF[6]  := INT_TO_STRING(debug_ID,'%d');
      LOG_MSG();
    END_IF;*)
    (*########################################################################*)

  END_IF;
ELSE
  DELAY_STOP := TX;  (* timer starten              *)
END_IF;
(*++++++++++++++++++++++++++++++++++++++++++++++++++++++++++++++++++++++++++*)

(* -----------------------------------------------------------------*)
(* wenn ein satelliten-baustein die portnummer 0 oder IP-Adresse    *)
(* 0.0.0.0 verwendet, sollen die am ip_control angegebene daten     *)
(* verwendet werden.           										*)
(* -----------------------------------------------------------------*)
IF IP_C.C_PORT = WORD#00 THEN
	IP_C.C_PORT := PORT; (* uebergebenen PORT durch paramtrierte PORT ersetzen *)
END_IF;
IF IP_C.C_IP=DWORD#00 AND IP_C.C_MODE<BYTE#4 THEN
	IP_C.C_IP := IP; (* uebergebene IP durch paramtrierte IP ersetzen *)
END_IF;

(* neue Verbindungs erwünscht ? *)
NEW_CONNECTION := C_IP <> IP_C.C_IP OR C_MODE <> IP_C.C_MODE OR C_PORT <> IP_C.C_PORT;

(* -----------------------------------------------------------------*)
(* Verbindungsparameter ausbereiten                                 *)
(* -----------------------------------------------------------------*)
IF IP_C.C_ENABLE AND NOT C_READY AND NEW_CONNECTION THEN

  (* neue Verbindungsparameter übernehmen *)
  C_IP   := IP_C.C_IP;
  C_MODE := IP_C.C_MODE;
  C_PORT := IP_C.C_PORT;

  (* -----------------------------------------------------------------*)
  (* CONNECTION_STRING erzeugen                                       *)
  (* Beispiel: '/UDP /ACTIVE /PORT=1000 /IP=192.168.178.1'            *)
  (*                                                                  *)
  (* Mode:                                                            *)
  (*  0: TCP + ACTIVE  + PORT + IP                                    *)
  (*  1: UDP + ACTIVE  + PORT + IP                                    *)
  (*  2: TCP + PASSIVE + PORT + IP                                    *)
  (*  3: UDP + PASSIVE + PORT + IP                                    *)
  (*  4: TCP + PASSIVE + PORT                                         *)
  (*  5: UDP + PASSIVE + PORT                                         *)
  (* -----------------------------------------------------------------*)

  (* bei allen ungeraden MODE Nummern UDP-String vorgeben *)
  CS := SEL_STRING((C_MODE AND BYTE#1) = BYTE#1,'','/UDP ');
  (* ACTIVE oder PASSIVE String anhängen *)
  CS := CONCAT(CS,SEL_STRING(C_MODE<BYTE#2,'/PASSIVE','/ACTIVE'));
  (* Portnummer String anhängen *)
  CS := CONCAT(CS,' /PORT=');
  CS := CONCAT(CS,WORD_TO_STRING(C_PORT,'%u'));

  IF C_MODE<BYTE#4 THEN
    IP4_TO_STRING(IP4:=C_IP);  (* String mit IP erzeugen *)
    CS := CONCAT(CS,' /IP=');
    CS := CONCAT(CS,IP4_TO_STRING.IP4_TO_STRING);
  END_IF;

  (*-------------------------------------------------------------------*)

  (* uebergebenen Timeout-Wert auf min-wert begrenzen *)
  ERROR_TIME := MAX(UDINT#200,TIME_TO_UDINT(TIME_OUT));
  IP_C.TIME_RESET := TRUE;   (* Alle Timer ruecksetzen *)

  (*####################  DEBUG-MESSAGE  ###################################*)
  (*IF _debug_enable THEN
    LOG_CL.NEW_MSG := 'IP_CON: ~1 -IP_ID ~6';
    LOG_CL.PRINTF[1] := CS;
    LOG_CL.PRINTF[6] := INT_TO_STRING(debug_ID,'%d');
    LOG_MSG();
  END_IF;*)
  (*########################################################################*)
END_IF;

(*++++++++++++++++++++++++++++++++++++++++++++++++++++++++++++++++++++++++++*)

C_ENABLE := IP_C.C_ENABLE AND NOT C_RECONNECT AND NOT NEW_CONNECTION AND IP_C.ERROR = DWORD#0;

(* -----------------------------------------------------------------*)
(* Systembaustein IP_CONNECT                                        *)
(* -----------------------------------------------------------------*)
FB_IP_CONNECT.EN_C    := C_ENABLE;
FB_IP_CONNECT.PARTNER := CS;
FB_IP_CONNECT();
C_READY  := FB_IP_CONNECT.VALID;
C_ERROR  := FB_IP_CONNECT.ERROR;
C_STATUS := FB_IP_CONNECT.STATUS;
C_ID     := FB_IP_CONNECT.ID;

(*++++++++++++++++++++++++++++++++++++++++++++++++++++++++++++++++++++++++++*)

IF C_ENABLE THEN
  IF NOT C_ENABLE_OLD THEN
    DELAY_VALUE := UDINT#50;  (* verzoegerungzeit vorgeben                     *)
    (*####################  DEBUG-MESSAGE  ###################################*)
    (*IF _debug_enable THEN
      LOG_CL.NEW_MSG := 'IP_CON: ENABLE + CYLCE-DELAY -IP_ID ~6';
      LOG_CL.PRINTF[6] := INT_TO_STRING(debug_ID,'%d');
      LOG_MSG();
    END_IF;*)
    (*########################################################################*)
  END_IF;
ELSE
  IF C_ENABLE_OLD THEN
    C_RECONNECT := FALSE;
    DELAY_VALUE := UDINT#50; (* verzoegerungzeit vorgeben                         *)
    (*####################  DEBUG-MESSAGE  ###################################*)
    (*IF _debug_enable THEN
      LOG_CL.NEW_MSG := 'IP_CON: DISABLE + CYLCE-DELAY -IP_ID ~6';
      LOG_CL.PRINTF[6] := INT_TO_STRING(debug_ID,'%d');
      LOG_MSG();
    END_IF;*)
    (*########################################################################*)
  END_IF;
END_IF;

C_ENABLE_OLD := C_ENABLE;

(*++++++++++++++++++++++++++++++++++++++++++++++++++++++++++++++++++++++++++*)

IF C_READY THEN
  IF NOT C_READY_OLD THEN
    (* Verbindung aufgebaut - positive Flanke erkannt*)
    IP_C.C_STATE := BYTE#254;
    DELAY_VALUE := UDINT#50;  (* verzoegerungzeit vorgeben *)
    IP_C.TIME_RESET := TRUE;  (* Alle Timer ruecksetzen *)
    (*####################  DEBUG-MESSAGE  ###################################*)
    (*IF _debug_enable THEN
      LOG_CL.NEW_MSG := 'IP_CON: CONNECTED -IP_ID ~6';
      LOG_CL.PRINTF[6] := INT_TO_STRING(debug_ID,'%d');
      LOG_MSG();
    END_IF;*)
    (*########################################################################*)
  ELSE
    IP_C.C_STATE := BYTE#255;  (* Verbindung ist aufgebaut                      *)
  END_IF;
ELSE
  IF C_READY_OLD THEN
    (* Verbindung abgebaut - negative Flanke erkannt*)
    IP_C.C_STATE := BYTE#1;
	IP_C.MAILBOX[1] := BYTE#0; (* Receive Info rücksetzen *)
	IP_C.MAILBOX[2] := BYTE#0; (* Send-Pause rücksetzen *)
	IP_C.MAILBOX[3] := BYTE#0; (* Receive-Pause rücksetzen *)
    DELAY_VALUE := UDINT#50;  (* verzoegerungzeit vorgeben *)

    IF NOT NEW_CONNECTION THEN
      S_ACTIVE := FALSE;        (* Sendeaktivitäten stoppen *)
      S_BUF.SIZE := UINT#0;     (* Sendelänge löschen       *)
      (*IP_C.TIME_RESET := TRUE;*)  (* Alle Timer ruecksetzen   *)
    END_IF;
    (*####################  DEBUG-MESSAGE  ###################################*)
    (*IF _debug_enable THEN
      LOG_CL.NEW_MSG := 'IP_CON: DISCONNECTED';
      LOG_MSG();
    END_IF;*)
    (*########################################################################*)
  ELSE
    IP_C.C_STATE := BYTE#000; (* Verbindung ist abgebaut *)
  END_IF;
END_IF;

C_READY_OLD := C_READY;
(*@KEY@: END_WORKSHEET *)
(*@KEY@: WORKSHEET
NAME: SEND
IEC_LANGUAGE: ST
*)
C := 1; (* voreinstellung: USEND nur einmal durchlaufen *)
IF S_BUF.SIZE > UINT#0 THEN
  IF C_READY AND C_ENABLE AND S_ACTIVE = FALSE AND IP_C.MAILBOX[2] = BYTE#0 THEN
    S_ACTIVE := TRUE; (* Sende-Betrieb aktivieren *)
    S_TIME := tx; (* Send Timer ruecksetzen *)
    R_TIME := tx; (* Receive Timer ruecksetzen *)
    C := 0; (* USEND zweimal aufrufen zur erzeugung einer positiven Flanke *)
    (*####################  DEBUG-MESSAGE  ###################################*)
    (*IF _debug_enable THEN
      LOG_CL.NEW_MSG := 'IP_SEN INIT: TOTAL: ~1 -IP_ID ~6';
      LOG_CL.PRINTF[1] := UINT_TO_STRING(S_BUF.SIZE,'%u');
      LOG_CL.PRINTF[6] := INT_TO_STRING(debug_ID,'%d');
      LOG_MSG();
    END_IF;*)
    (*########################################################################*)
  END_IF;
END_IF;

(* -----------------------------------------------------------------*)
(* Systembaustein IP_USEND (Datensenden)                            *)
(* -----------------------------------------------------------------*)
FOR C2 := C TO 1 DO
  FB_IP_USEND.REQ    := S_ACTIVE AND C2=1;
  FB_IP_USEND.ID     := C_ID;
  FB_IP_USEND.R_ID   := '';
  FB_IP_USEND.SD_1   := S_BUF;
  FB_IP_USEND();
  S_DONE   := FB_IP_USEND.DONE;
  S_ERROR  := FB_IP_USEND.ERROR;
  S_STATUS := FB_IP_USEND.STATUS;
  S_BUF    := FB_IP_USEND.SD_1;
END_FOR;

IF S_DONE THEN (* Daten fertig übertragen *)
    S_ACTIVE := FALSE;
    S_BUF.SIZE := UINT#0;
    (*####################  DEBUG-MESSAGE  ###################################*)
    (*IF _debug_enable THEN
      LOG_CL.NEW_MSG := 'IP_SEN FINISH -IP_ID ~6';
      LOG_CL.PRINTF[6] := INT_TO_STRING(debug_ID,'%d');
      LOG_MSG();
    END_IF;*)
    (*########################################################################*)

END_IF;

(*@KEY@: END_WORKSHEET *)
(*@KEY@: WORKSHEET
NAME: RECEIVE
IEC_LANGUAGE: ST
*)
(* -----------------------------------------------------------------*)
(* Systembaustein IP_URCV (Datenempfang)                            *)
(* -----------------------------------------------------------------*)

(* Die Empfangsbereitschaft wird zurückgenommen solange ein Sendevorgang läuft *)
(* sonst kann es vorkommen das die Antwort-daten schon empfangen werden,       *)
(* bevor der Sendevorgang vom programm abgeschlossen wurde *)

FB_IP_URCV.EN_R := C_READY AND NOT S_ACTIVE AND IP_C.MAILBOX[3] = BYTE#0;
FB_IP_URCV.ID   := C_ID;
FB_IP_URCV.R_ID := '';
FB_IP_URCV.RD_1 := R_BUF;
FB_IP_URCV();
R_NDR    := FB_IP_URCV.NDR;
R_ERROR  := FB_IP_URCV.ERROR;
R_STATUS := FB_IP_URCV.STATUS;
R_BUF    := FB_IP_URCV.RD_1;

(* -----------------------------------------------------------------*)
(* positive Flanke für Daten Empfangen abfragen                     *)
(* -----------------------------------------------------------------*)
IF R_NDR THEN
  	R_TIME := TX; (* Receive Timer ruecksetzen           *)
  	(* R_BUF.SIZE wird vom Empfangsbaustein automatisch beschrieben *)
    IP_C.MAILBOX[1] := USINT_TO_BYTE(BYTE_TO_USINT(IP_C.MAILBOX[1]) + USINT#1); (* Receive Info *)
    IF IP_C.MAILBOX[1] = BYTE#0 THEN IP_C.MAILBOX[1] := BYTE#1; END_IF;
    (*####################  DEBUG-MESSAGE  ###################################*)
    (*IF _debug_enable THEN
      LOG_CL.NEW_MSG := 'IP_REC DATA: SIZE: ~2 -IP_ID ~6';
      LOG_CL.PRINTF[2] := UINT_TO_STRING(R_BUF.SIZE,'%u');
      LOG_CL.PRINTF[6] := INT_TO_STRING(debug_ID,'%d');
      LOG_MSG();
    END_IF;*)
    (*########################################################################*)
END_IF;
(*@KEY@: END_WORKSHEET *)
(*@KEY@: WORKSHEET
NAME: ERROR
IEC_LANGUAGE: ST
*)
(* ----------------------------------------------------------------------------*)
(* Timer bearbeitung                                                           *)
(* ----------------------------------------------------------------------------*)
IF IP_C.TIME_RESET THEN     (* Alle Timer ruecksetzen      *)
  IP_C.TIME_RESET := FALSE; (* Reset rücksetzen            *)
  C_RECONNECT_COUNT := 0;   (* Reconnect zähler rücksetzen *)
  C_TIME := tx;             (* Connect   Timer ruecksetzen *)
  S_TIME := tx;             (* Send      Timer ruecksetzen *)
  R_TIME := tx;             (* Receive   Timer ruecksetzen *)

  ERROR_CON := BYTE#0;		(* Error Connect rücksetzen    *)
  ERROR_SND := BYTE#0;		(* Error Send rücksetzen       *)
  ERROR_RCV := BYTE#0;		(* Error Receive rücksetzen    *)
END_IF;

IF IP_C.R_OBSERVE = FALSE OR s_active THEN
    R_TIME := tx;
END_IF;

C_RECONNECT := FALSE;

(* ----------------------------------------------------------------------------*)
(* Error bearbeitung                                                           *)
(*                                                                             *)
(* bei pcworx ist nur wenn error = 1  der wert von status ein echter fehler    *)
(* status bekommt bei error "0" auch manchmal andere werte                     *)
(* ----------------------------------------------------------------------------*)

(* CONNECT Fehlercodes *)
IF ERROR_CON = BYTE#0 THEN
  IF C_ERROR THEN (* Die Verbindung wurde abgebrochen ignorieren *)
	IF C_STATUS = 16#31 THEN (* Die Verbindung wurde abgebrochen *)
		ERROR_CON := BYTE#253;
	ELSE
		ERROR_CON := INT_TO_BYTE(C_STATUS);
	END_IF;
  ELSIF TX - C_TIME > ERROR_TIME AND C_ENABLE AND NOT C_READY AND C_MODE < BYTE#2 THEN (* Connect Timeout *)
    IF C_RECONNECT_COUNT >= 3 THEN
      ERROR_CON := BYTE#255; (* Timeout-Fehler ausgeben *)
    ELSE
      C_TIME := TX; (* Connect   Timer ruecksetzen            *)
      C_RECONNECT_COUNT := C_RECONNECT_COUNT + 1;
      C_RECONNECT := TRUE;
      (*####################  DEBUG-MESSAGE  ###################################*)
      (*IF _debug_enable THEN
        LOG_CL.NEW_MSG := 'IP_CON: RECONNECT -IP_ID ~6';
        LOG_CL.PRINTF[6] := INT_TO_STRING(debug_ID,'%d');
        LOG_MSG();
      END_IF;*)
      (*########################################################################*)
    END_IF;
  END_IF;
END_IF;

(* SEND Fehlercodes *)
IF ERROR_SND = BYTE#0 THEN
  IF S_ERROR AND S_STATUS <> 16#65 THEN (* andere Bausteininstanz arbeitet mit dieser Verbindung *)
  	ERROR_SND := INT_TO_BYTE(S_STATUS);
  ELSIF TX - S_TIME > ERROR_TIME AND S_ACTIVE THEN (* Send Timeout *)
    ERROR_SND := BYTE#255; (* Timeout-Fehler ausgeben *)
  END_IF;
END_IF;

(* RECEIVE Fehlercodes *)
IF ERROR_RCV = BYTE#0 THEN
  IF R_ERROR AND (R_STATUS <> 16#33) AND (R_STATUS <> 16#31) AND (R_STATUS <> 16#65) THEN (* Receive Timeout,Verbindungsabbruch,andere Bausteininstanz arbeitet mit dieser Verbindung, ignorieren *)
  	ERROR_RCV := INT_TO_BYTE(R_STATUS);
  ELSIF TX - R_TIME > ERROR_TIME AND C_READY AND IP_C.R_OBSERVE THEN (* Receive Timeout *)
    ERROR_RCV := BYTE#255; (* Timeout-Fehler ausgeben *)
  END_IF;
END_IF;

IP_C.ERROR := DWORD_OF_BYTE(ERROR_CON,ERROR_SND,ERROR_RCV,BYTE#0);

(*####################  DEBUG-MESSAGE  ###################################*)
(*IF _debug_enable THEN
  IF (debug_last_id <> debug_ID) AND (IP_C.ERROR <> debug_lasterror) AND (IP_C.ERROR <> DWORD#00) THEN
    LOG_CL.NEW_MSG := 'IP_ERROR ~1 -IP_ID ~6';
    LOG_CL.PRINTF[1] := DWORD_TO_STRING(IP_C.ERROR,'%08X');
    LOG_CL.PRINTF[6] := INT_TO_STRING(debug_ID,'%d');
    LOG_MSG();
	debug_lasterror := IP_C.ERROR;
	debug_last_id   := debug_ID;
  END_IF;
END_IF;*)
(*########################################################################*)

(* revision history
ks	18. oct. 2008	rev 1.0
	original version
ks	05. jan. 2009	rev 1.1
	zusätzlichen Parameter "Port" hinzugefügt, und Code bei Verbindungsaufbau angepasst
ks	28. feb. 2009	rev 1.2
	connect code angepasst und verkürzung der zyklen bei Send
ks	20. oct. 2009	rev 1.3
	network_buffer basis 0
ks	06. dec. 2009	rev 1.4
	receive_count MAILBOX[1]
ks	10. nov. 2010	rev 1.5
	send_pause MAILBOX[2] and receive_pause MAILBOX[3]
ks	07. feb. 2011	rev 1.6
	Fehlercode 253 bei Remote-Verbindungsabbruch
ks	30. may. 2011	rev 1.7
	Fehler bei Empfangüberwachung
ks	26. jul. 2011	rev 1.8
	optimierung der Empfangsüberwachung
*)

(*@KEY@: END_WORKSHEET *)
END_FUNCTION_BLOCK

(* ---- LOG_VIEWPORT.ST ---- *)
(*@PROPERTIES_EX@
TYPE: POU
LOCALE: 0
IEC_LANGUAGE: ST
PLC_TYPE: independent
PROC_TYPE: independent
GROUP: NETWORK
*)
(*@KEY@:DESCRIPTION*)
(*
version 1.0		01 mai 2010
programmer		ks
tested BY		ks

LOG_VIEWPORT erzeugt einen Liste der Meldungen des Loggingbuffers die innerhalb einer virtuellen Ansicht enthalten sind.
*)

(*@KEY@:END_DESCRIPTION*)
FUNCTION_BLOCK LOG_VIEWPORT

(*Group:Parameter*)

VAR_IN_OUT
	LC :	us_LOG_CONTROL_80;
	LV :	us_LOG_VIEWPORT;
END_VAR

(*Group:lokal*)

VAR
	pos :	INT;
	count :	INT;
	idx :	INT;
	base :	INT;
	update_pos :	BOOL;
END_VAR

(*@KEY@: WORKSHEET
NAME: LOG_VIEWPORT
IEC_LANGUAGE: ST
*)
(* Scroll Button verarbeiten *)
IF LV.MOVE_TO_X <> 0 THEN
  CASE LV.MOVE_TO_X OF
  30000:
    pos := 1 ; (* älteste Meldung anzeigen *)
  30001:
    pos := LC.SIZE; (* neueste Meldung anzeigen *)
  30002:
    pos := pos + LV.COUNT; (* eine Seite nach unten blättern -> Richtung neuere Nachrichten *)
  30003:
    pos := pos - LV.COUNT; (* eine Seite nach oben blättern -> Richtung ältere Nachrichten *)
  ELSE
    pos := pos + LV.MOVE_TO_X;
  END_CASE;
  update_pos := TRUE;
  LV.MOVE_TO_X := 0;
END_IF;

IF (LV.UPDATE_COUNT <> LC.UPDATE_COUNT) OR update_pos THEN (* Aktualisierung überwachen *)
  LV.UPDATE := TRUE;
  LV.UPDATE_COUNT := LC.UPDATE_COUNT;
  update_pos := FALSE;

  (*-----------------------------------------------------------------------------------*)
  (* pos prüfen und übernehmen *)
  IF LC.RING_MODE THEN
    pos := LIMIT(1,pos,LC.SIZE - LV.COUNT + 1);
  ELSE
    IF LC.IDX > LV.COUNT THEN
      pos := LIMIT(1,pos,LC.IDX - LV.COUNT + 1);
    ELSE
      pos := 1;
    END_IF;
  END_IF;

  (*-----------------------------------------------------------------------------------*)
  (* idxBasis berechnen *)
  base := LC.IDX - pos - LV.COUNT + 1;
  IF LC.RING_MODE THEN
    (* Anzeige im Ringpuffermodus *)
    FOR count:= 1 TO LV.COUNT DO
      idx := base + count;
      IF idx < 1 THEN
        idx := idx + LC.SIZE;
      END_IF;
    END_FOR;
  ELSE
    (* Anzeige im Normalmodus *)
    FOR count:= 1 TO LV.COUNT DO
      idx := base + count;
      IF idx < 1 THEN
        (* Leere Zeile ausgeben *)
        LV.LINE_ARRAY[count] := 0;
      ELSE
        LV.LINE_ARRAY[count] := idx;
      END_IF;
    END_FOR;
  END_IF;
END_IF;

(* revision history
ks	01. mai 2010	rev 1.0
	original version
*)

(*@KEY@: END_WORKSHEET *)
END_FUNCTION_BLOCK

(* ---- MB_CLIENT.ST ---- *)
(*@PROPERTIES_EX@
TYPE: POU
LOCALE: 0
IEC_LANGUAGE: ST
PLC_TYPE: independent
PROC_TYPE: independent
GROUP: NETWORK
*)
(*@KEY@:DESCRIPTION*)

version 1.2		20. oct. 2009
programmer 		ks
tested by		ks

MB_CLIENT ermöglicht das Lesen/Schreiben von Daten über das Protokoll Modbus over Ethernet (OpenModbus)
(*@KEY@:END_DESCRIPTION*)
FUNCTION_BLOCK MB_CLIENT

(*Group:Default*)

VAR_IN_OUT
	IP_C :	oscat_IP_C;
	S_BUF :	oscat_NETWORK_BUFFER_SHORT;
	R_BUF :	oscat_NETWORK_BUFFER_SHORT;
	DATA :	oscat_aW0_255;
END_VAR

VAR_INPUT
	DATA_SIZE :	INT;
	ENABLE :	BOOL;
	UDP :	BOOL;
	FC :	INT;
	UNIT_ID :	BYTE;(*For Gateways only Slaveaddress*)
	R_ADDR :	INT;
	R_POINTS :	INT;
	R_DATA_ADR :	INT;
	R_DATA_BITPOS :	INT;
	W_ADDR :	INT;
	W_POINTS :	INT;
	W_DATA_ADR :	INT;
	W_DATA_BITPOS :	INT;
	DELAY :	TIME;
END_VAR

VAR_OUTPUT
	ERROR :	DWORD;
	BUSY :	BOOL;
END_VAR

VAR
	IP_STATE :	BYTE;
	IP_ID :	BYTE;
	IP_FIFO :	IP_FIFO;
	mask :	DWORD;
	w_tmp :	WORD;
	idx1 :	INT;
	idx2 :	INT;
	stop :	INT;
	i :	INT;
	bit_pos :	INT;
	w_mask :	WORD;
	b_mask :	BYTE;
	count :	INT;
	state :	INT;
	Transaction_ID :	INT;
	Response :	INT;
	comp :	INT;
	TON_1 :	TON;
END_VAR

(*@KEY@: WORKSHEET
NAME: MB_CLIENT
IEC_LANGUAGE: ST
*)

CASE state OF

00: (* Warten auf Delay-Time *)
	TON_1(IN:=ENABLE,PT:=DELAY);

  	IF TON_1.Q OR DELAY = T#0s THEN
		TON_1(IN:=FALSE);
		state := 20;
		IP_STATE := BYTE#1; (* Anmelden *)
	END_IF;

20: (* Bei IP_Control anmelden *)
	IF IP_STATE = BYTE#3 THEN
		(* IP Datenverkehr einrichten *)
		IP_C.C_PORT     := WORD#0;				(* Port von IP_CONTROL verwenden           		*)
		IP_C.C_IP       := DWORD#0;				(* IP von IP_CONTROL verwenden					*)
		IP_C.C_MODE     := BOOL_TO_BYTE(UDP);	(* Mode: 0=TCP+ACTIVE+IP , 1=UDP+ACTIVE+IP   	*)
		IP_C.TIME_RESET := TRUE;				(* Zeitueberwachung rücksetzen                  *)
		IP_C.C_ENABLE   := TRUE;				(* Verbindungsaufbau freigeben                  *)
		IP_C.R_OBSERVE  := TRUE;				(* Empfangsueberwachung                         *)

		(******************************************************************)
		ERROR := DWORD#00; (* letzten Fehler rücksetzen *)

		CASE FC OF

		(******************************************************************)
		1..2: (* 0x01 Read Coil Status , 0x02 Read Input Status *)
			IF R_POINTS <= 2000 THEN
				w_tmp := INT_TO_WORD(R_ADDR);
				S_BUF.BUFFER[08] := WORD_TO_BYTE(SHR(w_tmp,8));
				S_BUF.BUFFER[09] := WORD_TO_BYTE(w_tmp);
				w_tmp := INT_TO_WORD(R_POINTS);
				S_BUF.BUFFER[10] := WORD_TO_BYTE(SHR(w_tmp,8));
				S_BUF.BUFFER[11] := WORD_TO_BYTE(w_tmp);
				S_BUF.SIZE := UINT#12;
				Response :=	WORD_TO_INT(SHR(INT_TO_WORD(R_POINTS + 7),3));
				comp := 7;
			ELSE
				ERROR := DWORD#2; (* ILLEGAL DATA ADDRESS *)
			END_IF;
		(******************************************************************)
		3..4: (* 0x03 Read Holding Registers , 0x04 Read Input Registers *)
			IF R_POINTS <= 125 THEN
				w_tmp := INT_TO_WORD(R_ADDR);
				S_BUF.BUFFER[08] := WORD_TO_BYTE(SHR(w_tmp,8));
				S_BUF.BUFFER[09] := WORD_TO_BYTE(w_tmp);
				w_tmp := INT_TO_WORD(R_POINTS);
				S_BUF.BUFFER[10] := WORD_TO_BYTE(SHR(w_tmp,8));
				S_BUF.BUFFER[11] := WORD_TO_BYTE(w_tmp);

				S_BUF.SIZE := UINT#12;
				Response :=	WORD_TO_INT(SHL(w_tmp,1));
				comp := 7;
			ELSE
				ERROR := DWORD#2; (* ILLEGAL DATA ADDRESS *)
			END_IF;
		(******************************************************************)
		5:	(* 0x05 Force Single Coil *)
			IF W_DATA_ADR <= DATA_SIZE THEN
				w_tmp := INT_TO_WORD(W_ADDR);
				S_BUF.BUFFER[08] := WORD_TO_BYTE(SHR(w_tmp,8));
				S_BUF.BUFFER[09] := WORD_TO_BYTE(w_tmp);
				S_BUF.BUFFER[10] := SEL((DATA[W_DATA_ADR] AND SHL(WORD#1,W_DATA_BITPOS))>WORD#00,BYTE#16#00,BYTE#16#FF);
				S_BUF.BUFFER[11] := BYTE#00;

				S_BUF.SIZE := UINT#12;
				Response :=	3;
				comp := 11;
			ELSE
				ERROR := DWORD#2; (* ILLEGAL DATA ADDRESS *)
			END_IF;
		(******************************************************************)
		6:	(* 0x06 Preset Single Register *)
			IF W_DATA_ADR <= DATA_SIZE THEN
				w_tmp := INT_TO_WORD(W_ADDR);
				S_BUF.BUFFER[08] := WORD_TO_BYTE(SHR(w_tmp,8));
				S_BUF.BUFFER[09] := WORD_TO_BYTE(w_tmp);
				w_tmp := DATA[W_DATA_ADR];
				S_BUF.BUFFER[10] := WORD_TO_BYTE(SHR(w_tmp,8));
				S_BUF.BUFFER[11] := WORD_TO_BYTE(w_tmp);

				S_BUF.SIZE := UINT#12;
				Response :=	3;
				comp := 11;
			ELSE
				ERROR := DWORD#2; (* ILLEGAL DATA ADDRESS *)
			END_IF;
		(******************************************************************)
		15:	(* 0x0F Force Multiple Coils *)
			IF (WORD_TO_INT(SHR(INT_TO_WORD(WORD_TO_INT(SHL(INT_TO_WORD(W_DATA_ADR),4)) + W_POINTS + W_DATA_BITPOS + 15),4)) <= DATA_SIZE) AND W_POINTS <= 1968 THEN
				w_tmp := INT_TO_WORD(W_ADDR);
				S_BUF.BUFFER[08] := WORD_TO_BYTE(SHR(w_tmp,8));
				S_BUF.BUFFER[09] := WORD_TO_BYTE(w_tmp);
				w_tmp := INT_TO_WORD(W_POINTS);
				S_BUF.BUFFER[10] := WORD_TO_BYTE(SHR(w_tmp,8));
				S_BUF.BUFFER[11] := WORD_TO_BYTE(w_tmp);
				S_BUF.BUFFER[12] := WORD_TO_BYTE(SHR(INT_TO_WORD(W_POINTS + 7),3));

				w_mask := SHL(WORD#1,W_DATA_BITPOS);
				bit_pos := 0;
				w_tmp := WORD#00;
				idx1 := 12;
				idx2 := W_DATA_ADR;
				FOR i := 1 TO W_POINTS DO
					w_tmp :=BIT_LOAD_W(w_tmp,(DATA[idx2] AND w_mask)>WORD#0,bit_pos);
					bit_pos := bit_pos + 1;
					IF bit_pos > 7 OR i=W_POINTS THEN
						bit_pos := 0;
						idx1 := idx1 + 1;
						S_BUF.BUFFER[idx1] := WORD_TO_BYTE(w_tmp);
						w_tmp := WORD#0;
					END_IF;
					w_mask := ROL(w_mask,1);
					IF w_mask = WORD#1 THEN
						idx2 := idx2 + 1;
					END_IF;
				END_FOR;
				S_BUF.SIZE := INT_TO_UINT(idx1+1);
				Response :=	3;
				comp := 11;
			ELSE
				ERROR := DWORD#2; (* ILLEGAL DATA ADDRESS *)
			END_IF;
		(******************************************************************)
		16:	(* 0x10 Write Multiple Registers *)
			IF W_DATA_ADR + W_POINTS <= DATA_SIZE AND W_POINTS <= 123 THEN
				w_tmp := INT_TO_WORD(W_ADDR);
				S_BUF.BUFFER[08] := WORD_TO_BYTE(SHR(w_tmp,8));
				S_BUF.BUFFER[09] := WORD_TO_BYTE(w_tmp);
				w_tmp := INT_TO_WORD(W_POINTS);
				S_BUF.BUFFER[10] := WORD_TO_BYTE(SHR(w_tmp,8));
				S_BUF.BUFFER[11] := WORD_TO_BYTE(w_tmp);
				S_BUF.BUFFER[12] := SHL(S_BUF.BUFFER[11],1);

				idx1 := 11;
				count := W_DATA_ADR + W_POINTS - 1;
				FOR i := W_DATA_ADR TO count DO
					idx1 := idx1 + 2;
					idx2 := idx1 + 1; (* zweiter index für pcworx notwendig ! *)
					w_tmp := DATA[i];
					S_BUF.BUFFER[idx1] := WORD_TO_BYTE(SHR(w_tmp,8));
					S_BUF.BUFFER[idx2] := WORD_TO_BYTE(w_tmp);
				END_FOR;

				S_BUF.SIZE := INT_TO_UINT(idx2 + 1);
				Response := 3;
				comp := 11;
			ELSE
				ERROR := DWORD#2; (* ILLEGAL DATA ADDRESS *)
			END_IF;
		(******************************************************************)
		22:	(* 0x16 Mask Write Register *)
			IF W_DATA_ADR + 2 <= DATA_SIZE THEN
				w_tmp := INT_TO_WORD(W_ADDR);
				S_BUF.BUFFER[08] := WORD_TO_BYTE(SHR(w_tmp,8));
				S_BUF.BUFFER[09] := WORD_TO_BYTE(w_tmp);
				idx1 := W_DATA_ADR;
				w_tmp := DATA[idx1];
				S_BUF.BUFFER[10] := WORD_TO_BYTE(SHR(w_tmp,8));
				S_BUF.BUFFER[11] := WORD_TO_BYTE(w_tmp);
				idx1 := idx1 +1;
				w_tmp := DATA[idx1];
				S_BUF.BUFFER[12] := WORD_TO_BYTE(SHR(w_tmp,8));
				S_BUF.BUFFER[13] := WORD_TO_BYTE(w_tmp);

				S_BUF.SIZE := UINT#14;
				Response :=	5;
				comp := 13;
			ELSE
				ERROR := DWORD#2; (* ILLEGAL DATA ADDRESS *)
			END_IF;
		(******************************************************************)
		23:	(* 0x17 Read/Write Multible Registers *)
			IF W_DATA_ADR + W_POINTS <= DATA_SIZE AND W_POINTS <= 121 AND R_POINTS <= 125 THEN
				idx1 := 15;
				count := W_DATA_ADR + W_POINTS - 1;
				FOR i := W_DATA_ADR TO count DO
					idx1 := idx1 + 2;
					idx2 := idx1 + 1; (* zweiter index für pcworx notwendig ! *)
					w_tmp := DATA[i];
					S_BUF.BUFFER[idx1] := WORD_TO_BYTE(SHR(w_tmp,8));
					S_BUF.BUFFER[idx2] := WORD_TO_BYTE(w_tmp);
				END_FOR;

				(* WRITE *)
				w_tmp := INT_TO_WORD(W_ADDR);
				S_BUF.BUFFER[12] := WORD_TO_BYTE(SHR(w_tmp,8));
				S_BUF.BUFFER[13] := WORD_TO_BYTE(w_tmp);
				w_tmp := INT_TO_WORD(W_POINTS);
				S_BUF.BUFFER[14] := WORD_TO_BYTE(SHR(w_tmp,8));
				S_BUF.BUFFER[15] := WORD_TO_BYTE(w_tmp);
				S_BUF.BUFFER[16] := SHL(S_BUF.BUFFER[15],1);

				(* READ *)
				w_tmp := INT_TO_WORD(R_ADDR);
				S_BUF.BUFFER[08] := WORD_TO_BYTE(SHR(w_tmp,8));
				S_BUF.BUFFER[09] := WORD_TO_BYTE(w_tmp);
				w_tmp := INT_TO_WORD(R_POINTS);
				S_BUF.BUFFER[10] := WORD_TO_BYTE(SHR(w_tmp,8));
				S_BUF.BUFFER[11] := WORD_TO_BYTE(w_tmp);

				S_BUF.SIZE := INT_TO_UINT(idx2+1);
				Response :=	WORD_TO_INT(SHL(w_tmp,1));
				comp := 7;
			ELSE
				ERROR := DWORD#2; (* ILLEGAL DATA ADDRESS *)
			END_IF;
		(******************************************************************)

		ELSE
			ERROR := DWORD#00000001;	(* ILLEGAL FUNCTION *)
		END_CASE;

		(* Daten senden *)
		IF ERROR = DWORD#00 THEN
			Transaction_ID := Transaction_ID + 1;
			w_tmp := UINT_TO_WORD(S_BUF.SIZE - UINT#6);
			(* ---- H E A D E R --------------------------------------------------------------- *)
			S_BUF.BUFFER[0] := IP_ID;								(* TRANSACTION-ID HI-Byte 	*)
			S_BUF.BUFFER[1] := INT_TO_BYTE(Transaction_ID);			(* TRANSACTION-ID LO-Byte	*)
			S_BUF.BUFFER[2] := BYTE#00;								(* PROTOKOLL-ID HI-Byte 	*)
			S_BUF.BUFFER[3] := BYTE#00;								(* PROTOKOLL-ID LO-Byte 	*)
			S_BUF.BUFFER[4] := WORD_TO_BYTE(SHR(w_tmp,8));			(* Laenge HI-Byte			*)
			S_BUF.BUFFER[5] := WORD_TO_BYTE(w_tmp);					(* Laenge LO-Byte			*)
			S_BUF.BUFFER[6] := UNIT_ID;								(* UNIT						*)
			S_BUF.BUFFER[7] := INT_TO_BYTE(FC);						(* FUNCTION-CODE			*)
			(*----- END OF HEADER --------------------------------------------------------------*)
			R_BUF.SIZE := UINT#0; (* Empfangsbuffer löschen *)
			state := 30; (* wait for response *)
		ELSE
			IP_STATE := BYTE#4; (* Abmelden *)
			state := 00;
		END_IF;
	END_IF;

30: (* response *)
	IF IP_C.ERROR <> DWORD#00 THEN
    	ERROR := IP_C.ERROR;
		IP_STATE := BYTE#4; (* Abmelden *)
		state := 00;

	ELSIF S_BUF.SIZE = UINT#0 AND R_BUF.SIZE > UINT#0 THEN

		(* erwartete länge in sendebuffer nachträglich eintragen um vergleich zu ermöglichen *)
		w_tmp := INT_TO_WORD(Response + 3);
		S_BUF.BUFFER[4] := WORD_TO_BYTE(SHR(w_tmp,8));
		S_BUF.BUFFER[5] := WORD_TO_BYTE(w_tmp);

		FOR i := 0 TO comp DO
			IF S_BUF.BUFFER[i] <> R_BUF.BUFFER[i] THEN EXIT; END_IF;
		END_FOR;

		IF R_BUF.SIZE >= UINT#9 AND R_BUF.BUFFER[7] > BYTE#128 THEN  (* Bit 7 = Error Message *)
			ERROR := BYTE_TO_DWORD(R_BUF.BUFFER[8]);
			IP_STATE := BYTE#4; (* Abmelden *)
			state := 00;

		ELSIF R_BUF.SIZE = INT_TO_UINT(Response + 9) AND i > comp THEN
			mask := SHL(DWORD#1,FC);

			(* READ_COILS, READ_INPUT_DISCRETES *)
			IF (mask AND DWORD#2#00000000_00000000_00000000_00000110) <> DWORD#0 THEN (* FC 1,2 *)
				IF WORD_TO_INT(SHR(INT_TO_WORD(WORD_TO_INT(SHL(INT_TO_WORD(R_DATA_ADR),4)) + R_POINTS + R_DATA_BITPOS + 15),4)) <= DATA_SIZE THEN
					b_mask := BYTE#1;
					idx1 := 09;
					idx2 := R_DATA_ADR;
					bit_pos := R_DATA_BITPOS;
					FOR i := 1 TO R_POINTS DO
						DATA[idx2]:=BIT_LOAD_W(DATA[idx2],(R_BUF.BUFFER[idx1] AND b_mask)>BYTE#0,bit_pos);
						bit_pos := bit_pos + 1;
						IF bit_pos > 15 THEN
							idx2 := idx2 + 1;
							bit_pos := 0;
						END_IF;
						b_mask := ROL(b_mask,1);
						IF b_mask = BYTE#1 THEN
							idx1 := idx1 +1;
						END_IF;
					END_FOR;
				ELSE
					ERROR := DWORD#2; (* ILLEGAL DATA ADDRESS *)
				END_IF;

			(* READ_MULTIPLE_REGISTERS, READ_INPUT_REGISTERS, READ_WRITE_REGISTERS *)
			ELSIF (mask AND DWORD#2#00000000_10000000_00000000_00011000) <> DWORD#0 THEN (* FC 3,4,23 *)
				IF R_DATA_ADR + R_POINTS <= DATA_SIZE THEN
					stop := R_DATA_ADR + R_POINTS -1 ;
					idx1 := 07;
					FOR i := R_DATA_ADR TO stop DO
						idx1 := idx1 +2;
						idx2 := idx1 +1;
						DATA[i] := WORD_OF_BYTE(R_BUF.BUFFER[idx1],R_BUF.BUFFER[idx2]);
					END_FOR;
				ELSE
					ERROR := DWORD#2; (* ILLEGAL DATA ADDRESS *)
				END_IF;
			ELSIF (mask AND DWORD#2#11111111_00111110_01111111_10000001) > DWORD#0 THEN (* ILLEGAL FUNCTION CODE ? *)
				ERROR := DWORD#1; (* ILLEGAL FUNCTION *)
			END_IF;
		ELSE
			ERROR := DWORD#3; (* ILLEGAL DATA VALUE *)
		END_IF;

		IP_STATE := BYTE#4; (* Abmelden *)
		state := 00;
		R_BUF.SIZE := UINT#0;

	END_IF;

END_CASE;

(* IP_FIFO *)
IP_FIFO(FIFO:=IP_C.FIFO,STATE:=IP_STATE,ID:=IP_ID);
IP_C.FIFO:=IP_FIFO.FIFO;
IP_STATE := IP_FIFO.STATE;
IP_ID:=IP_FIFO.ID;

BUSY := IP_STATE = BYTE#3;

(* revision history
ks	05. jan. 2009	rev 1.0
	original version

ks	28. jan. 2009	rev 1.1
	network_buffer_short verwendet

ks	20. oct. 2009	rev 1.2
Networkbuffer und Buffer-funktionen auf Basis 0

*)
(*@KEY@: END_WORKSHEET *)
END_FUNCTION_BLOCK

(* ---- MB_SERVER.ST ---- *)
(*@PROPERTIES_EX@
TYPE: POU
LOCALE: 0
IEC_LANGUAGE: ST
PLC_TYPE: independent
PROC_TYPE: independent
GROUP: NETWORK
*)
(*@KEY@:DESCRIPTION*)
version 1.3		17. may. 2011
programmer 		ks
tested by		ks

MB_SERVER ermöglicht das Lesen/Schreiben von Daten durch ein Remote-Device mittels Modbus over Ethernet (OpenModbus)
(*@KEY@:END_DESCRIPTION*)
FUNCTION_BLOCK MB_SERVER

(*Group:Default*)

VAR_IN_OUT
	IP_C :	oscat_IP_C;
	S_BUF :	oscat_NETWORK_BUFFER_SHORT;
	R_BUF :	oscat_NETWORK_BUFFER_SHORT;
	VMAP :	oscat_MB_VMAP;
	DATA :	oscat_aW0_255;
END_VAR

VAR_INPUT
	DATA_SIZE :	INT;
	ENABLE :	BOOL;
	UDP :	BOOL;
END_VAR

VAR_OUTPUT
	ERROR :	DWORD;
END_VAR

VAR
	MB_VMAP :	MB_VMAP;
	adr1 :	INT;
	adr2 :	INT;
	points :	INT;
	points2 :	INT;
	coils :	BYTE;
	mask :	BYTE;
	idx1 :	INT;
	idx2 :	INT;
	bit_pos :	INT;
	count :	INT;
	fc :	INT;
	i :	INT;
	state :	INT;
	IP_STATE :	BYTE;
	IP_ID :	BYTE;
	IP_FIFO :	IP_FIFO;
	w_tmp :	WORD;
	last_cycle :	TIME;
	tx :	TIME;
	T_PLC_MS :	T_PLC_MS;
	t :	TON;
	ip_error :	BOOL;
END_VAR

(*@KEY@: WORKSHEET
NAME: MB_SERVER
IEC_LANGUAGE: ST
*)
(* read system time *)
T_PLC_MS();
tx := UDINT_TO_TIME(T_PLC_MS.T_PLC_MS);

FOR i := 1 TO 10 DO
	IF VMAP[i].TIME_OUT > T#0s THEN
		VMAP[i].TIME_OUT := VMAP[i].TIME_OUT + tx - last_cycle;
	END_IF;
END_FOR;
last_cycle := tx;
ip_error := IP_C.ERROR > DWORD#0;

CASE state OF

00: (* Warten auf Freigabe *)
  	IF ENABLE THEN
		state := 10;
		IP_STATE := BYTE#1; (* Anmelden *)
	END_IF;

10: (* Bei IP_Control anmelden und auf freigabe warten *)
	IF IP_STATE = BYTE#3 THEN

  		(* IP Datenverkehr einrichten *)
		IP_C.C_PORT     := WORD#0;					(* Port von IP_CONTROL verwenden           		 *)
  		IP_C.C_IP       := DWORD#0;					(* IP von IP_CONTROL verwenden					 *)
  		IP_C.C_MODE     := SEL(UDP,BYTE#4,BYTE#5);	(* Mode: 4=TCP+PASSIV+PORT , 5=UDP+PASSIV+PORT   *)
  		IP_C.TIME_RESET := TRUE;					(* Zeitueberwachung rücksetzen                   *)
  		IP_C.C_ENABLE   := TRUE;					(* Verbindungsaufbau freigeben                   *)
  		IP_C.R_OBSERVE  := FALSE;					(* keine Empfangsueberwachung                    *)
  		state := 20;
	END_IF;

20:	IF NOT ip_error THEN
	 	IF S_BUF.SIZE = UINT#0 AND R_BUF.SIZE > UINT#6 THEN	(* Datensenden nicht aktiv und Daten wurden empfangen *)
			IF  R_BUF.SIZE = WORD_TO_UINT(WORD_OF_BYTE(R_BUF.BUFFER[4],R_BUF.BUFFER[5])) + UINT#6 THEN (* gültige Datenlänge *)
				ERROR := DWORD#00;	 (* Error löschen *)

				(* Header kopieren *)
				FOR i := 0 TO 13 DO
					S_BUF.BUFFER[i] := R_BUF.BUFFER[i];
				END_FOR;

				fc := _BYTE_TO_INT(R_BUF.BUFFER[7]);

				adr1 := WORD_TO_INT(WORD_OF_BYTE(R_BUF.BUFFER[8],R_BUF.BUFFER[9]));
				points := WORD_TO_INT(WORD_OF_BYTE(R_BUF.BUFFER[10],R_BUF.BUFFER[11]));

				(* Virtual Address *)
				MB_VMAP(VMAP:=VMAP,FC:=fc,V_ADR:=adr1,V_CNT:=points,SIZE:=DATA_SIZE);
				VMAP:=MB_VMAP.VMAP;
				adr1:=MB_VMAP.P_ADR;
				bit_pos:=MB_VMAP.P_BIT;
				ERROR:=BYTE_TO_DWORD(MB_VMAP.ERROR);

				IF ERROR = DWORD#0 THEN
					CASE fc OF

					(*--------------------------------------------------*)
					1..2 : (* Read Coil Status / Read Input Status 		*)
						count := 9; (* erstes Datenbyte *)
						coils := BYTE#0;
						mask := BYTE#1;
						FOR i := 1 TO points DO
							IF mask = BYTE#0 THEN
								mask := BYTE#1;
								S_BUF.BUFFER[count] := coils;
								coils := BYTE#0;
								count := count + 1;
							END_IF;
							IF (DATA[adr1] AND SHL(WORD#1,bit_pos)) > WORD#0 THEN
								coils := coils OR mask;
							END_IF;

							bit_Pos := bit_Pos + 1;
							IF bit_pos > 15 THEN
								adr1 := adr1 + 1;
								bit_pos := 0;
							END_IF;

							mask := SHL(mask,1);
						END_FOR;
						S_BUF.BUFFER[Count] := coils;

						S_BUF.BUFFER[8] := INT_TO_BYTE(count - 8);  (* Bytecount *)
						S_BUF.SIZE := INT_TO_UINT(count + 1);

					(*--------------------------------------------------*)
					3..4 : (* Read Holding Registers / Read Input Registers *)
						idx1 := 07;
						count := adr1 + points - 1;
						FOR i := adr1 TO count DO
							idx1 := idx1 + 2;
							idx2 := idx1 + 1; (* zweiter index für pcworx notwendig ! *)
							w_tmp := DATA[i];
							S_BUF.BUFFER[idx1] := WORD_TO_BYTE(SHR(w_tmp,8));
							S_BUF.BUFFER[idx2] := WORD_TO_BYTE(w_tmp);
						END_FOR;
						S_BUF.BUFFER[8] := SHL(INT_TO_BYTE(points),1); (* Anzahl Register in Bytes *)
						S_BUF.SIZE := INT_TO_UINT(idx2 + 1);
					(*--------------------------------------------------*)
					5 : (* Force Single Coil *)
						DATA[adr1]:=BIT_LOAD_W(DATA[adr1],R_BUF.BUFFER[10]>BYTE#0,bit_pos);
						S_BUF.SIZE := UINT#12;
					(*--------------------------------------------------*)
					6 : (* Preset Single Register *)
						DATA[adr1] := WORD_OF_BYTE(R_BUF.BUFFER[10],R_BUF.BUFFER[11]);
						S_BUF.SIZE := UINT#12;
					(*--------------------------------------------------*)
					15 : (* Force Multible Coils *)
						mask := BYTE#1;
						idx1 := 13;
						FOR i := 1 TO points DO
							DATA[adr1]:=BIT_LOAD_W(DATA[adr1],(R_BUF.BUFFER[idx1] AND mask)>BYTE#0,bit_pos);
							bit_pos := bit_pos + 1;
							IF bit_pos > 15 THEN
								adr1 := adr1 + 1;
								bit_pos := 0;
							END_IF;
							mask := ROL(mask,1);
							IF mask = BYTE#1 THEN
								idx1 := idx1 +1;
							END_IF;
						END_FOR;
						S_BUF.SIZE := UINT#12;
					(*--------------------------------------------------*)
					16 : (* Preset Multiple Registers	*)
						idx1 := 11;
						count := adr1 + points -1;
						FOR i := adr1 TO Count DO
							idx1 := idx1 + 2;
	 						idx2 := idx1 + 1;
							Data[i] := WORD_OF_BYTE(R_BUF.BUFFER[idx1],R_BUF.BUFFER[idx2]);
						END_FOR;
						S_BUF.SIZE := UINT#12;
					(*--------------------------------------------------*)
					22 : (* Mask Write Register *)
						w_tmp := WORD_OF_BYTE(R_BUF.BUFFER[11],R_BUF.BUFFER[11]); (* and mask *)
						DATA[adr1] := (DATA[adr1] AND w_tmp) OR (WORD_OF_BYTE(R_BUF.BUFFER[12],R_BUF.BUFFER[13]) AND (NOT w_tmp));
						S_BUF.SIZE := UINT#14;
					(*--------------------------------------------------*)
					23 : (* Read / Write Registers	*)
						(*--- Write-Register -----------------------------------*)
						adr2 := WORD_TO_INT(WORD_OF_BYTE(R_BUF.BUFFER[12],R_BUF.BUFFER[13]));
						points2 := WORD_TO_INT(WORD_OF_BYTE(R_BUF.BUFFER[14],R_BUF.BUFFER[15]));

						(* Virtual Address Write Register *)
						MB_VMAP(VMAP:=VMAP,FC:=16,V_ADR:=adr2,V_CNT:=points2,SIZE:=DATA_SIZE);
						VMAP:=MB_VMAP.VMAP;
						adr2:=MB_VMAP.P_ADR;
						ERROR:=BYTE_TO_DWORD(MB_VMAP.ERROR);

						IF ERROR = DWORD#0 THEN
							idx1 := 15;
							count := adr2 + points2 -1;
							FOR i := adr2 TO count DO
								idx1 := idx1 + 2;
	 							idx2 := idx1 + 1; (* zweiter index für pcworx notwendig ! *)
								Data[i] := WORD_OF_BYTE(R_BUF.BUFFER[idx1],R_BUF.BUFFER[idx2]);
							END_FOR;

							(*--- Read-Register -----------------------------------*)
							idx1 := 07;
							count := adr1 + points - 1;
							FOR i := adr1 TO count DO
								idx1 := idx1 + 2;
								idx2 := idx1 + 1; (* zweiter index für pcworx notwendig ! *)
								w_tmp := DATA[i];
								S_BUF.BUFFER[idx1] := WORD_TO_BYTE(SHR(w_tmp,8));
								S_BUF.BUFFER[idx2] := WORD_TO_BYTE(w_tmp);
							END_FOR;
							S_BUF.BUFFER[8] := SHL(INT_TO_BYTE(points),1); (* Anzahl Register in Bytes *)
							S_BUF.SIZE := INT_TO_UINT(idx2 + 1);

						END_IF;

					(*--------------------------------------------------*)
					ELSE
						ERROR := DWORD#01; (* ILLEGAL FUNCTION *)
					END_CASE;
				END_IF;
			END_IF;

			IF ERROR > DWORD#0 THEN
				S_BUF.BUFFER[7] := S_BUF.BUFFER[7] OR BYTE#2#1000_0000; (* Fehlerbit setzen *)
				S_BUF.BUFFER[8] := DWORD_TO_BYTE(ERROR);
				S_BUF.SIZE := UINT#9;
			END_IF;

			S_BUF.BUFFER[4] := BYTE#0; (* high Byte *)
			S_BUF.BUFFER[5] := UINT_TO_BYTE(S_BUF.SIZE - UINT#6); (* Längenfeld eintragen - nur low byte *)

		END_IF;
	ELSE
		ERROR := IP_C.ERROR;
	END_IF;

	t(IN:= ip_error, PT:=T#5s);
	IF t.Q THEN
		IP_C.TIME_RESET := TRUE; (* Error Reset *)
	END_IF;

	R_BUF.SIZE := UINT#0; (* Empfangsdaten zerstören *)

	IF ENABLE = FALSE THEN
	    IP_STATE := BYTE#4; (* Abmelden *)
		state := 00;
	END_IF;
END_CASE;

(* IP_FIFO *)
IP_FIFO(FIFO:=IP_C.FIFO,STATE:=IP_STATE,ID:=IP_ID);
IP_C.FIFO:=IP_FIFO.FIFO;
IP_STATE := IP_FIFO.STATE;
IP_ID:=IP_FIFO.ID;

(* revision history
ks	05. jan. 2009	rev 1.0
	original version

ks	28. jan. 2009	rev 1.1
	network_buffer_short verwendet

ks	20. oct. 2009	rev 1.2
	change lokal-var adr to adr1,Networkbuffer und Buffer-funktionen auf Basis 0

ks	17. may. 2011	rev 1.3
	automatischer re-connect
*)

(*@KEY@: END_WORKSHEET *)
END_FUNCTION_BLOCK
